//     PlcTask Outputs/GVL_iXlinker.Device_1_EtherCAT.Term_1_EK1200.Term_2_EL6002.COM_RxPDO_Map_Outputs_Channel_1.Data_Out[3] <-> COM RxPDO-Map Outputs Channel 1/Data Out 3
//     PlcTask Outputs/GVL_iXlinker.Device_1_EtherCAT.Term_1_EK1200.Term_2_EL6002.COM_RxPDO_Map_Outputs_Channel_1.Data_Out[4] <-> COM RxPDO-Map Outputs Channel 1/Data Out 4
//     PlcTask Outputs/GVL_iXlinker.Device_1_EtherCAT.Term_1_EK1200.Term_2_EL6002.COM_RxPDO_Map_Outputs_Channel_1.Data_Out[5] <-> COM RxPDO-Map Outputs Channel 1/Data Out 5
//     PlcTask Outputs/GVL_iXlinker.Device_1_EtherCAT.Term_1_EK1200.Term_2_EL6002.COM_RxPDO_Map_Outputs_Channel_1.Data_Out[6] <-> COM RxPDO-Map Outputs Channel 1/Data Out 6
//     PlcTask Outputs/GVL_iXlinker.Device_1_EtherCAT.Term_1_EK1200.Term_2_EL6002.COM_RxPDO_Map_Outputs_Channel_1.Data_Out[7] <-> COM RxPDO-Map Outputs Channel 1/Data Out 7
//     PlcTask Outputs/GVL_iXlinker.Device_1_EtherCAT.Term_1_EK1200.Term_2_EL6002.COM_RxPDO_Map_Outputs_Channel_1.Data_Out[8] <-> COM RxPDO-Map Outputs Channel 1/Data Out 8
//     PlcTask Outputs/GVL_iXlinker.Device_1_EtherCAT.Term_1_EK1200.Term_2_EL6002.COM_RxPDO_Map_Outputs_Channel_1.Data_Out[9] <-> COM RxPDO-Map Outputs Channel 1/Data Out 9
//     PlcTask Outputs/GVL_iXlinker.Device_1_EtherCAT.Term_1_EK1200.Term_2_EL6002.COM_RxPDO_Map_Outputs_Channel_2.Data_Out[0] <-> COM RxPDO-Map Outputs Channel 2/Data Out 0
//     PlcTask Outputs/GVL_iXlinker.Device_1_EtherCAT.Term_1_EK1200.Term_2_EL6002.COM_RxPDO_Map_Outputs_Channel_2.Data_Out[10] <-> COM RxPDO-Map Outputs Channel 2/Data Out 10
//     PlcTask Outputs/GVL_iXlinker.Device_1_EtherCAT.Term_1_EK1200.Term_2_EL6002.COM_RxPDO_Map_Outputs_Channel_2.Data_Out[11] <-> COM RxPDO-Map Outputs Channel 2/Data Out 11
//     PlcTask Outputs/GVL_iXlinker.Device_1_EtherCAT.Term_1_EK1200.Term_2_EL6002.COM_RxPDO_Map_Outputs_Channel_2.Data_Out[12] <-> COM RxPDO-Map Outputs Channel 2/Data Out 12
//     PlcTask Outputs/GVL_iXlinker.Device_1_EtherCAT.Term_1_EK1200.Term_2_EL6002.COM_RxPDO_Map_Outputs_Channel_2.Data_Out[13] <-> COM RxPDO-Map Outputs Channel 2/Data Out 13
//     PlcTask Outputs/GVL_iXlinker.Device_1_EtherCAT.Term_1_EK1200.Term_2_EL6002.COM_RxPDO_Map_Outputs_Channel_2.Data_Out[14] <-> COM RxPDO-Map Outputs Channel 2/Data Out 14
//     PlcTask Outputs/GVL_iXlinker.Device_1_EtherCAT.Term_1_EK1200.Term_2_EL6002.COM_RxPDO_Map_Outputs_Channel_2.Data_Out[15] <-> COM RxPDO-Map Outputs Channel 2/Data Out 15
//     PlcTask Outputs/GVL_iXlinker.Device_1_EtherCAT.Term_1_EK1200.Term_2_EL6002.COM_RxPDO_Map_Outputs_Channel_2.Data_Out[16] <-> COM RxPDO-Map Outputs Channel 2/Data Out 16
//     PlcTask Outputs/GVL_iXlinker.Device_1_EtherCAT.Term_1_EK1200.Term_2_EL6002.COM_RxPDO_Map_Outputs_Channel_2.Data_Out[17] <-> COM RxPDO-Map Outputs Channel 2/Data Out 17
//     PlcTask Outputs/GVL_iXlinker.Device_1_EtherCAT.Term_1_EK1200.Term_2_EL6002.COM_RxPDO_Map_Outputs_Channel_2.Data_Out[18] <-> COM RxPDO-Map Outputs Channel 2/Data Out 18
//     PlcTask Outputs/GVL_iXlinker.Device_1_EtherCAT.Term_1_EK1200.Term_2_EL6002.COM_RxPDO_Map_Outputs_Channel_2.Data_Out[19] <-> COM RxPDO-Map Outputs Channel 2/Data Out 19
//     PlcTask Outputs/GVL_iXlinker.Device_1_EtherCAT.Term_1_EK1200.Term_2_EL6002.COM_RxPDO_Map_Outputs_Channel_2.Data_Out[1] <-> COM RxPDO-Map Outputs Channel 2/Data Out 1
//     PlcTask Outputs/GVL_iXlinker.Device_1_EtherCAT.Term_1_EK1200.Term_2_EL6002.COM_RxPDO_Map_Outputs_Channel_2.Data_Out[20] <-> COM RxPDO-Map Outputs Channel 2/Data Out 20
//     PlcTask Outputs/GVL_iXlinker.Device_1_EtherCAT.Term_1_EK1200.Term_2_EL6002.COM_RxPDO_Map_Outputs_Channel_2.Data_Out[21] <-> COM RxPDO-Map Outputs Channel 2/Data Out 21
//     PlcTask Outputs/GVL_iXlinker.Device_1_EtherCAT.Term_1_EK1200.Term_2_EL6002.COM_RxPDO_Map_Outputs_Channel_2.Data_Out[2] <-> COM RxPDO-Map Outputs Channel 2/Data Out 2
//     PlcTask Outputs/GVL_iXlinker.Device_1_EtherCAT.Term_1_EK1200.Term_2_EL6002.COM_RxPDO_Map_Outputs_Channel_2.Data_Out[3] <-> COM RxPDO-Map Outputs Channel 2/Data Out 3
//     PlcTask Outputs/GVL_iXlinker.Device_1_EtherCAT.Term_1_EK1200.Term_2_EL6002.COM_RxPDO_Map_Outputs_Channel_2.Data_Out[4] <-> COM RxPDO-Map Outputs Channel 2/Data Out 4
//     PlcTask Outputs/GVL_iXlinker.Device_1_EtherCAT.Term_1_EK1200.Term_2_EL6002.COM_RxPDO_Map_Outputs_Channel_2.Data_Out[5] <-> COM RxPDO-Map Outputs Channel 2/Data Out 5
//     PlcTask Outputs/GVL_iXlinker.Device_1_EtherCAT.Term_1_EK1200.Term_2_EL6002.COM_RxPDO_Map_Outputs_Channel_2.Data_Out[6] <-> COM RxPDO-Map Outputs Channel 2/Data Out 6
//     PlcTask Outputs/GVL_iXlinker.Device_1_EtherCAT.Term_1_EK1200.Term_2_EL6002.COM_RxPDO_Map_Outputs_Channel_2.Data_Out[7] <-> COM RxPDO-Map Outputs Channel 2/Data Out 7
//     PlcTask Outputs/GVL_iXlinker.Device_1_EtherCAT.Term_1_EK1200.Term_2_EL6002.COM_RxPDO_Map_Outputs_Channel_2.Data_Out[8] <-> COM RxPDO-Map Outputs Channel 2/Data Out 8
//     PlcTask Outputs/GVL_iXlinker.Device_1_EtherCAT.Term_1_EK1200.Term_2_EL6002.COM_RxPDO_Map_Outputs_Channel_2.Data_Out[9] <-> COM RxPDO-Map Outputs Channel 2/Data Out 9
//   TcoIoTests/TcoIoTests Instance <-> Device 1 (EtherCAT)/Term 1 (EK1200)/Term 3 (EL1809)
//     PlcTask Inputs/GVL_iXlinker.Device_1_EtherCAT.Term_1_EK1200.Term_3_EL1809.Channel_{1..16}.Input <-> Channel {1..16}/Input  (16 links)
//     PlcTask Inputs/GVL_iXlinker.Device_1_EtherCAT.Term_1_EK1200.Term_3_EL1809.InfoData.State <-> InfoData/State
//     PlcTask Inputs/GVL_iXlinker.Device_1_EtherCAT.Term_1_EK1200.Term_3_EL1809.WcState.InputToggle <-> WcState/InputToggle
//     PlcTask Inputs/GVL_iXlinker.Device_1_EtherCAT.Term_1_EK1200.Term_3_EL1809.WcState.WcState <-> WcState/WcState
//   TcoIoTests/TcoIoTests Instance <-> Device 1 (EtherCAT)/Term 1 (EK1200)/Term 4 (EL2809)
//     PlcTask Inputs/GVL_iXlinker.Device_1_EtherCAT.Term_1_EK1200.Term_4_EL2809.InfoData.State <-> InfoData/State
//     PlcTask Inputs/GVL_iXlinker.Device_1_EtherCAT.Term_1_EK1200.Term_4_EL2809.WcState.WcState <-> WcState/WcState
//     PlcTask Outputs/GVL_iXlinker.Device_1_EtherCAT.Term_1_EK1200.Term_4_EL2809.Channel_{1..16}.Output <-> Channel {1..16}/Output  (16 links)
//   TcoIoTests/TcoIoTests Instance <-> Device 1 (EtherCAT)/Term 1 (EK1200)/Term 5 (EL4004)
//     PlcTask Inputs/GVL_iXlinker.Device_1_EtherCAT.Term_1_EK1200.Term_5_EL4004.InfoData.AdsAddr <-> InfoData/AdsAddr
//     PlcTask Inputs/GVL_iXlinker.Device_1_EtherCAT.Term_1_EK1200.Term_5_EL4004.InfoData.State <-> InfoData/State
//     PlcTask Inputs/GVL_iXlinker.Device_1_EtherCAT.Term_1_EK1200.Term_5_EL4004.WcState.WcState <-> WcState/WcState
//     PlcTask Outputs/GVL_iXlinker.Device_1_EtherCAT.Term_1_EK1200.Term_5_EL4004.AO_Outputs_Channel_{1..4}.Analog_output <-> AO Outputs Channel {1..4}/Analog output  (4 links)
//   TcoIoTests/TcoIoTests Instance <-> Device 1 (EtherCAT)/Term 1 (EK1200)/Term 6 (EL2809)
//     PlcTask Inputs/GVL_iXlinker.Device_1_EtherCAT.Term_1_EK1200.Term_6_EL2809.InfoData.State <-> InfoData/State
//     PlcTask Inputs/GVL_iXlinker.Device_1_EtherCAT.Term_1_EK1200.Term_6_EL2809.WcState.WcState <-> WcState/WcState
//     PlcTask Outputs/GVL_iXlinker.Device_1_EtherCAT.Term_1_EK1200.Term_6_EL2809.Channel_{1..16}.Output <-> Channel {1..16}/Output  (16 links)
//   TcoIoTests/TcoIoTests Instance <-> Device 1 (EtherCAT)/Term 1 (EK1200)/Term 7 (EL6001)
//     PlcTask Inputs/GVL_iXlinker.Device_1_EtherCAT.Term_1_EK1200.Term_7_EL6001.COM_Inputs.Data_In[{0..21}] <-> COM Inputs/Data In {0..21}  (22 links)
//     PlcTask Inputs/GVL_iXlinker.Device_1_EtherCAT.Term_1_EK1200.Term_7_EL6001.COM_Inputs.Status/Buffer_full <-> COM Inputs/Status/Buffer full
//     PlcTask Inputs/GVL_iXlinker.Device_1_EtherCAT.Term_1_EK1200.Term_7_EL6001.COM_Inputs.Status/Framing_error <-> COM Inputs/Status/Framing error
//     PlcTask Inputs/GVL_iXlinker.Device_1_EtherCAT.Term_1_EK1200.Term_7_EL6001.COM_Inputs.Status/Init_accepted <-> COM Inputs/Status/Init accepted
//     PlcTask Inputs/GVL_iXlinker.Device_1_EtherCAT.Term_1_EK1200.Term_7_EL6001.COM_Inputs.Status/Input_length <-> COM Inputs/Status/Input length
//     PlcTask Inputs/GVL_iXlinker.Device_1_EtherCAT.Term_1_EK1200.Term_7_EL6001.COM_Inputs.Status/Overrun_error <-> COM Inputs/Status/Overrun error
//     PlcTask Inputs/GVL_iXlinker.Device_1_EtherCAT.Term_1_EK1200.Term_7_EL6001.COM_Inputs.Status/Parity_error <-> COM Inputs/Status/Parity error
//     PlcTask Inputs/GVL_iXlinker.Device_1_EtherCAT.Term_1_EK1200.Term_7_EL6001.COM_Inputs.Status/Receive_request <-> COM Inputs/Status/Receive request
//     PlcTask Inputs/GVL_iXlinker.Device_1_EtherCAT.Term_1_EK1200.Term_7_EL6001.COM_Inputs.Status/Transmit_accepted <-> COM Inputs/Status/Transmit accepted
//     PlcTask Inputs/GVL_iXlinker.Device_1_EtherCAT.Term_1_EK1200.Term_7_EL6001.InfoData.AdsAddr <-> InfoData/AdsAddr
//     PlcTask Inputs/GVL_iXlinker.Device_1_EtherCAT.Term_1_EK1200.Term_7_EL6001.InfoData.State <-> InfoData/State
//     PlcTask Inputs/GVL_iXlinker.Device_1_EtherCAT.Term_1_EK1200.Term_7_EL6001.WcState.InputToggle <-> WcState/InputToggle
//     PlcTask Inputs/GVL_iXlinker.Device_1_EtherCAT.Term_1_EK1200.Term_7_EL6001.WcState.WcState <-> WcState/WcState
//     PlcTask Outputs/GVL_iXlinker.Device_1_EtherCAT.Term_1_EK1200.Term_7_EL6001.COM_Outputs.Ctrl/Init_request <-> COM Outputs/Ctrl/Init request
//     PlcTask Outputs/GVL_iXlinker.Device_1_EtherCAT.Term_1_EK1200.Term_7_EL6001.COM_Outputs.Ctrl/Output_length <-> COM Outputs/Ctrl/Output length
//     PlcTask Outputs/GVL_iXlinker.Device_1_EtherCAT.Term_1_EK1200.Term_7_EL6001.COM_Outputs.Ctrl/Receive_accepted <-> COM Outputs/Ctrl/Receive accepted
//     PlcTask Outputs/GVL_iXlinker.Device_1_EtherCAT.Term_1_EK1200.Term_7_EL6001.COM_Outputs.Ctrl/Send_continues <-> COM Outputs/Ctrl/Send continues
//     PlcTask Outputs/GVL_iXlinker.Device_1_EtherCAT.Term_1_EK1200.Term_7_EL6001.COM_Outputs.Ctrl/Transmit_request <-> COM Outputs/Ctrl/Transmit request
//     PlcTask Outputs/GVL_iXlinker.Device_1_EtherCAT.Term_1_EK1200.Term_7_EL6001.COM_Outputs.Data_Out[{0..21}] <-> COM Outputs/Data Out {0..21}  (22 links)
//   TcoIoTests/TcoIoTests Instance <-> Device 2 (EtherCAT)
//     PlcTask Inputs/GVL_iXlinker.Device_2_EtherCAT.InfoData.AmsNetId <-> InfoData/AmsNetId
//     PlcTask Inputs/GVL_iXlinker.Device_2_EtherCAT.InfoData.CfgSlaveCount <-> InfoData/CfgSlaveCount
//     PlcTask Inputs/GVL_iXlinker.Device_2_EtherCAT.InfoData.ChangeCount <-> InfoData/ChangeCount
//     PlcTask Inputs/GVL_iXlinker.Device_2_EtherCAT.InfoData.DevId <-> InfoData/DevId
//     PlcTask Inputs/GVL_iXlinker.Device_2_EtherCAT.Inputs.DevState <-> Inputs/DevState
//     PlcTask Inputs/GVL_iXlinker.Device_2_EtherCAT.Inputs.Frm0InputToggle <-> Inputs/Frm0InputToggle
//     PlcTask Inputs/GVL_iXlinker.Device_2_EtherCAT.Inputs.Frm0State <-> Inputs/Frm0State
//     PlcTask Inputs/GVL_iXlinker.Device_2_EtherCAT.Inputs.Frm0WcState <-> Inputs/Frm0WcState
//     PlcTask Inputs/GVL_iXlinker.Device_2_EtherCAT.Inputs.SlaveCount <-> Inputs/SlaveCount
//     PlcTask Outputs/GVL_iXlinker.Device_2_EtherCAT.Outputs.DevCtrl <-> Outputs/DevCtrl
//     PlcTask Outputs/GVL_iXlinker.Device_2_EtherCAT.Outputs.Frm0Ctrl <-> Outputs/Frm0Ctrl
//     PlcTask Outputs/GVL_iXlinker.Device_2_EtherCAT.Outputs.Frm0WcCtrl <-> Outputs/Frm0WcCtrl
//   TcoIoTests/TcoIoTests Instance <-> Device 2 (EtherCAT)/Term 9 (EK1100)
//     PlcTask Inputs/GVL_iXlinker.Device_2_EtherCAT.Term_9_EK1100.InfoData.State <-> InfoData/State
//   TcoIoTests/TcoIoTests Instance <-> Device 2 (EtherCAT)/Term 9 (EK1100)/Term 10 (EK1122)
//     PlcTask Inputs/GVL_iXlinker.Device_2_EtherCAT.Term_9_EK1100.Term_10_EK1122.InfoData.State <-> InfoData/State
//   TcoIoTests/TcoIoTests Instance <-> Device 2 (EtherCAT)/Term 9 (EK1100)/Term 10 (EK1122)/Term 11 (EK1100)
//     PlcTask Inputs/GVL_iXlinker.Device_2_EtherCAT.Term_9_EK1100.Term_10_EK1122.Term_11_EK1100.InfoData.State <-> InfoData/State
//   TcoIoTests/TcoIoTests Instance <-> Device 2 (EtherCAT)/Term 9 (EK1100)/Term 10 (EK1122)/Term 11 (EK1100)/Term 12 (EL3174-0002)
//     PlcTask Inputs/GVL_iXlinker.Device_2_EtherCAT.Term_9_EK1100.Term_10_EK1122.Term_11_EK1100.Term_12_EL3174_0002.AI_Standard_Channel_1.Status/Error <-> AI Standard Channel 1/Status/Error
//     PlcTask Inputs/GVL_iXlinker.Device_2_EtherCAT.Term_9_EK1100.Term_10_EK1122.Term_11_EK1100.Term_12_EL3174_0002.AI_Standard_Channel_2.Status/Error <-> AI Standard Channel 2/Status/Error
//     PlcTask Inputs/GVL_iXlinker.Device_2_EtherCAT.Term_9_EK1100.Term_10_EK1122.Term_11_EK1100.Term_12_EL3174_0002.AI_Standard_Channel_3.Status/Error <-> AI Standard Channel 3/Status/Error
//     PlcTask Inputs/GVL_iXlinker.Device_2_EtherCAT.Term_9_EK1100.Term_10_EK1122.Term_11_EK1100.Term_12_EL3174_0002.AI_Standard_Channel_4.Status/Error <-> AI Standard Channel 4/Status/Error
//     PlcTask Inputs/GVL_iXlinker.Device_2_EtherCAT.Term_9_EK1100.Term_10_EK1122.Term_11_EK1100.Term_12_EL3174_0002.AI_Standard_Channel_1.Status/Limit_1 <-> AI Standard Channel 1/Status/Limit 1
//     PlcTask Inputs/GVL_iXlinker.Device_2_EtherCAT.Term_9_EK1100.Term_10_EK1122.Term_11_EK1100.Term_12_EL3174_0002.AI_Standard_Channel_1.Status/Limit_2 <-> AI Standard Channel 1/Status/Limit 2
//     PlcTask Inputs/GVL_iXlinker.Device_2_EtherCAT.Term_9_EK1100.Term_10_EK1122.Term_11_EK1100.Term_12_EL3174_0002.AI_Standard_Channel_2.Status/Limit_1 <-> AI Standard Channel 2/Status/Limit 1
//     PlcTask Inputs/GVL_iXlinker.Device_2_EtherCAT.Term_9_EK1100.Term_10_EK1122.Term_11_EK1100.Term_12_EL3174_0002.AI_Standard_Channel_2.Status/Limit_2 <-> AI Standard Channel 2/Status/Limit 2
//     PlcTask Inputs/GVL_iXlinker.Device_2_EtherCAT.Term_9_EK1100.Term_10_EK1122.Term_11_EK1100.Term_12_EL3174_0002.AI_Standard_Channel_3.Status/Limit_1 <-> AI Standard Channel 3/Status/Limit 1
//     PlcTask Inputs/GVL_iXlinker.Device_2_EtherCAT.Term_9_EK1100.Term_10_EK1122.Term_11_EK1100.Term_12_EL3174_0002.AI_Standard_Channel_3.Status/Limit_2 <-> AI Standard Channel 3/Status/Limit 2
//     PlcTask Inputs/GVL_iXlinker.Device_2_EtherCAT.Term_9_EK1100.Term_10_EK1122.Term_11_EK1100.Term_12_EL3174_0002.AI_Standard_Channel_4.Status/Limit_1 <-> AI Standard Channel 4/Status/Limit 1
//     PlcTask Inputs/GVL_iXlinker.Device_2_EtherCAT.Term_9_EK1100.Term_10_EK1122.Term_11_EK1100.Term_12_EL3174_0002.AI_Standard_Channel_4.Status/Limit_2 <-> AI Standard Channel 4/Status/Limit 2
//     PlcTask Inputs/GVL_iXlinker.Device_2_EtherCAT.Term_9_EK1100.Term_10_EK1122.Term_11_EK1100.Term_12_EL3174_0002.AI_Standard_Channel_1.Status/Overrange <-> AI Standard Channel 1/Status/Overrange
//     PlcTask Inputs/GVL_iXlinker.Device_2_EtherCAT.Term_9_EK1100.Term_10_EK1122.Term_11_EK1100.Term_12_EL3174_0002.AI_Standard_Channel_2.Status/Overrange <-> AI Standard Channel 2/Status/Overrange
//     PlcTask Inputs/GVL_iXlinker.Device_2_EtherCAT.Term_9_EK1100.Term_10_EK1122.Term_11_EK1100.Term_12_EL3174_0002.AI_Standard_Channel_3.Status/Overrange <-> AI Standard Channel 3/Status/Overrange
//     PlcTask Inputs/GVL_iXlinker.Device_2_EtherCAT.Term_9_EK1100.Term_10_EK1122.Term_11_EK1100.Term_12_EL3174_0002.AI_Standard_Channel_4.Status/Overrange <-> AI Standard Channel 4/Status/Overrange
//     PlcTask Inputs/GVL_iXlinker.Device_2_EtherCAT.Term_9_EK1100.Term_10_EK1122.Term_11_EK1100.Term_12_EL3174_0002.AI_Standard_Channel_1.Status/Sync_error <-> AI Standard Channel 1/Status/Sync error
//     PlcTask Inputs/GVL_iXlinker.Device_2_EtherCAT.Term_9_EK1100.Term_10_EK1122.Term_11_EK1100.Term_12_EL3174_0002.AI_Standard_Channel_2.Status/Sync_error <-> AI Standard Channel 2/Status/Sync error
//     PlcTask Inputs/GVL_iXlinker.Device_2_EtherCAT.Term_9_EK1100.Term_10_EK1122.Term_11_EK1100.Term_12_EL3174_0002.AI_Standard_Channel_3.Status/Sync_error <-> AI Standard Channel 3/Status/Sync error
//     PlcTask Inputs/GVL_iXlinker.Device_2_EtherCAT.Term_9_EK1100.Term_10_EK1122.Term_11_EK1100.Term_12_EL3174_0002.AI_Standard_Channel_4.Status/Sync_error <-> AI Standard Channel 4/Status/Sync error
//     PlcTask Inputs/GVL_iXlinker.Device_2_EtherCAT.Term_9_EK1100.Term_10_EK1122.Term_11_EK1100.Term_12_EL3174_0002.AI_Standard_Channel_1.Status/TxPDO_State <-> AI Standard Channel 1/Status/TxPDO State
//     PlcTask Inputs/GVL_iXlinker.Device_2_EtherCAT.Term_9_EK1100.Term_10_EK1122.Term_11_EK1100.Term_12_EL3174_0002.AI_Standard_Channel_2.Status/TxPDO_State <-> AI Standard Channel 2/Status/TxPDO State
//     PlcTask Inputs/GVL_iXlinker.Device_2_EtherCAT.Term_9_EK1100.Term_10_EK1122.Term_11_EK1100.Term_12_EL3174_0002.AI_Standard_Channel_3.Status/TxPDO_State <-> AI Standard Channel 3/Status/TxPDO State
//     PlcTask Inputs/GVL_iXlinker.Device_2_EtherCAT.Term_9_EK1100.Term_10_EK1122.Term_11_EK1100.Term_12_EL3174_0002.AI_Standard_Channel_4.Status/TxPDO_State <-> AI Standard Channel 4/Status/TxPDO State
//     PlcTask Inputs/GVL_iXlinker.Device_2_EtherCAT.Term_9_EK1100.Term_10_EK1122.Term_11_EK1100.Term_12_EL3174_0002.AI_Standard_Channel_1.Status/TxPDO_Toggle <-> AI Standard Channel 1/Status/TxPDO Toggle
//     PlcTask Inputs/GVL_iXlinker.Device_2_EtherCAT.Term_9_EK1100.Term_10_EK1122.Term_11_EK1100.Term_12_EL3174_0002.AI_Standard_Channel_2.Status/TxPDO_Toggle <-> AI Standard Channel 2/Status/TxPDO Toggle
//     PlcTask Inputs/GVL_iXlinker.Device_2_EtherCAT.Term_9_EK1100.Term_10_EK1122.Term_11_EK1100.Term_12_EL3174_0002.AI_Standard_Channel_3.Status/TxPDO_Toggle <-> AI Standard Channel 3/Status/TxPDO Toggle
//     PlcTask Inputs/GVL_iXlinker.Device_2_EtherCAT.Term_9_EK1100.Term_10_EK1122.Term_11_EK1100.Term_12_EL3174_0002.AI_Standard_Channel_4.Status/TxPDO_Toggle <-> AI Standard Channel 4/Status/TxPDO Toggle
//     PlcTask Inputs/GVL_iXlinker.Device_2_EtherCAT.Term_9_EK1100.Term_10_EK1122.Term_11_EK1100.Term_12_EL3174_0002.AI_Standard_Channel_1.Status/Underrange <-> AI Standard Channel 1/Status/Underrange
//     PlcTask Inputs/GVL_iXlinker.Device_2_EtherCAT.Term_9_EK1100.Term_10_EK1122.Term_11_EK1100.Term_12_EL3174_0002.AI_Standard_Channel_2.Status/Underrange <-> AI Standard Channel 2/Status/Underrange
//     PlcTask Inputs/GVL_iXlinker.Device_2_EtherCAT.Term_9_EK1100.Term_10_EK1122.Term_11_EK1100.Term_12_EL3174_0002.AI_Standard_Channel_3.Status/Underrange <-> AI Standard Channel 3/Status/Underrange
//     PlcTask Inputs/GVL_iXlinker.Device_2_EtherCAT.Term_9_EK1100.Term_10_EK1122.Term_11_EK1100.Term_12_EL3174_0002.AI_Standard_Channel_4.Status/Underrange <-> AI Standard Channel 4/Status/Underrange
//     PlcTask Inputs/GVL_iXlinker.Device_2_EtherCAT.Term_9_EK1100.Term_10_EK1122.Term_11_EK1100.Term_12_EL3174_0002.AI_Standard_Channel_1.Value <-> AI Standard Channel 1/Value
//     PlcTask Inputs/GVL_iXlinker.Device_2_EtherCAT.Term_9_EK1100.Term_10_EK1122.Term_11_EK1100.Term_12_EL3174_0002.AI_Standard_Channel_2.Value <-> AI Standard Channel 2/Value
//     PlcTask Inputs/GVL_iXlinker.Device_2_EtherCAT.Term_9_EK1100.Term_10_EK1122.Term_11_EK1100.Term_12_EL3174_0002.AI_Standard_Channel_3.Value <-> AI Standard Channel 3/Value
//     PlcTask Inputs/GVL_iXlinker.Device_2_EtherCAT.Term_9_EK1100.Term_10_EK1122.Term_11_EK1100.Term_12_EL3174_0002.AI_Standard_Channel_4.Value <-> AI Standard Channel 4/Value
//     PlcTask Inputs/GVL_iXlinker.Device_2_EtherCAT.Term_9_EK1100.Term_10_EK1122.Term_11_EK1100.Term_12_EL3174_0002.InfoData.AdsAddr <-> InfoData/AdsAddr
//     PlcTask Inputs/GVL_iXlinker.Device_2_EtherCAT.Term_9_EK1100.Term_10_EK1122.Term_11_EK1100.Term_12_EL3174_0002.InfoData.State <-> InfoData/State
//     PlcTask Inputs/GVL_iXlinker.Device_2_EtherCAT.Term_9_EK1100.Term_10_EK1122.Term_11_EK1100.Term_12_EL3174_0002.WcState.InputToggle <-> WcState/InputToggle
//     PlcTask Inputs/GVL_iXlinker.Device_2_EtherCAT.Term_9_EK1100.Term_10_EK1122.Term_11_EK1100.Term_12_EL3174_0002.WcState.WcState <-> WcState/WcState
//   TcoIoTests/TcoIoTests Instance <-> Device 2 (EtherCAT)/Term 9 (EK1100)/Term 10 (EK1122)/Term 11 (EK1100)/Term 13 (EL6001)
//     PlcTask Inputs/GVL_iXlinker.Device_2_EtherCAT.Term_9_EK1100.Term_10_EK1122.Term_11_EK1100.Term_13_EL6001.COM_Inputs.Data_In[{0..21}] <-> COM Inputs/Data In {0..21}  (22 links)
//     PlcTask Inputs/GVL_iXlinker.Device_2_EtherCAT.Term_9_EK1100.Term_10_EK1122.Term_11_EK1100.Term_13_EL6001.COM_Inputs.Status/Buffer_full <-> COM Inputs/Status/Buffer full
//     PlcTask Inputs/GVL_iXlinker.Device_2_EtherCAT.Term_9_EK1100.Term_10_EK1122.Term_11_EK1100.Term_13_EL6001.COM_Inputs.Status/Framing_error <-> COM Inputs/Status/Framing error
//     PlcTask Inputs/GVL_iXlinker.Device_2_EtherCAT.Term_9_EK1100.Term_10_EK1122.Term_11_EK1100.Term_13_EL6001.COM_Inputs.Status/Init_accepted <-> COM Inputs/Status/Init accepted
//     PlcTask Inputs/GVL_iXlinker.Device_2_EtherCAT.Term_9_EK1100.Term_10_EK1122.Term_11_EK1100.Term_13_EL6001.COM_Inputs.Status/Input_length <-> COM Inputs/Status/Input length
//     PlcTask Inputs/GVL_iXlinker.Device_2_EtherCAT.Term_9_EK1100.Term_10_EK1122.Term_11_EK1100.Term_13_EL6001.COM_Inputs.Status/Overrun_error <-> COM Inputs/Status/Overrun error
//     PlcTask Inputs/GVL_iXlinker.Device_2_EtherCAT.Term_9_EK1100.Term_10_EK1122.Term_11_EK1100.Term_13_EL6001.COM_Inputs.Status/Parity_error <-> COM Inputs/Status/Parity error
//     PlcTask Inputs/GVL_iXlinker.Device_2_EtherCAT.Term_9_EK1100.Term_10_EK1122.Term_11_EK1100.Term_13_EL6001.COM_Inputs.Status/Receive_request <-> COM Inputs/Status/Receive request
//     PlcTask Inputs/GVL_iXlinker.Device_2_EtherCAT.Term_9_EK1100.Term_10_EK1122.Term_11_EK1100.Term_13_EL6001.COM_Inputs.Status/Transmit_accepted <-> COM Inputs/Status/Transmit accepted
//     PlcTask Inputs/GVL_iXlinker.Device_2_EtherCAT.Term_9_EK1100.Term_10_EK1122.Term_11_EK1100.Term_13_EL6001.InfoData.AdsAddr <-> InfoData/AdsAddr
//     PlcTask Inputs/GVL_iXlinker.Device_2_EtherCAT.Term_9_EK1100.Term_10_EK1122.Term_11_EK1100.Term_13_EL6001.InfoData.State <-> InfoData/State
//     PlcTask Inputs/GVL_iXlinker.Device_2_EtherCAT.Term_9_EK1100.Term_10_EK1122.Term_11_EK1100.Term_13_EL6001.WcState.InputToggle <-> WcState/InputToggle
//     PlcTask Inputs/GVL_iXlinker.Device_2_EtherCAT.Term_9_EK1100.Term_10_EK1122.Term_11_EK1100.Term_13_EL6001.WcState.WcState <-> WcState/WcState
//     PlcTask Outputs/GVL_iXlinker.Device_2_EtherCAT.Term_9_EK1100.Term_10_EK1122.Term_11_EK1100.Term_13_EL6001.COM_Outputs.Ctrl/Init_request <-> COM Outputs/Ctrl/Init request
//     PlcTask Outputs/GVL_iXlinker.Device_2_EtherCAT.Term_9_EK1100.Term_10_EK1122.Term_11_EK1100.Term_13_EL6001.COM_Outputs.Ctrl/Output_length <-> COM Outputs/Ctrl/Output length
//     PlcTask Outputs/GVL_iXlinker.Device_2_EtherCAT.Term_9_EK1100.Term_10_EK1122.Term_11_EK1100.Term_13_EL6001.COM_Outputs.Ctrl/Receive_accepted <-> COM Outputs/Ctrl/Receive accepted
//     PlcTask Outputs/GVL_iXlinker.Device_2_EtherCAT.Term_9_EK1100.Term_10_EK1122.Term_11_EK1100.Term_13_EL6001.COM_Outputs.Ctrl/Send_continues <-> COM Outputs/Ctrl/Send continues
//     PlcTask Outputs/GVL_iXlinker.Device_2_EtherCAT.Term_9_EK1100.Term_10_EK1122.Term_11_EK1100.Term_13_EL6001.COM_Outputs.Ctrl/Transmit_request <-> COM Outputs/Ctrl/Transmit request
//     PlcTask Outputs/GVL_iXlinker.Device_2_EtherCAT.Term_9_EK1100.Term_10_EK1122.Term_11_EK1100.Term_13_EL6001.COM_Outputs.Data_Out[{0..21}] <-> COM Outputs/Data Out {0..21}  (22 links)
//   TcoIoTests/TcoIoTests Instance <-> Device 2 (EtherCAT)/Term 9 (EK1100)/Term 10 (EK1122)/Term 11 (EK1100)/Term 14 (EL3011)
//     PlcTask Inputs/GVL_iXlinker.Device_2_EtherCAT.Term_9_EK1100.Term_10_EK1122.Term_11_EK1100.Term_14_EL3011.AI_Standard.Status/Error <-> AI Standard/Status/Error
//     PlcTask Inputs/GVL_iXlinker.Device_2_EtherCAT.Term_9_EK1100.Term_10_EK1122.Term_11_EK1100.Term_14_EL3011.AI_Standard.Status/Limit_1 <-> AI Standard/Status/Limit 1
//     PlcTask Inputs/GVL_iXlinker.Device_2_EtherCAT.Term_9_EK1100.Term_10_EK1122.Term_11_EK1100.Term_14_EL3011.AI_Standard.Status/Limit_2 <-> AI Standard/Status/Limit 2
//     PlcTask Inputs/GVL_iXlinker.Device_2_EtherCAT.Term_9_EK1100.Term_10_EK1122.Term_11_EK1100.Term_14_EL3011.AI_Standard.Status/Overrange <-> AI Standard/Status/Overrange
//     PlcTask Inputs/GVL_iXlinker.Device_2_EtherCAT.Term_9_EK1100.Term_10_EK1122.Term_11_EK1100.Term_14_EL3011.AI_Standard.Status/TxPDO_State <-> AI Standard/Status/TxPDO State
//     PlcTask Inputs/GVL_iXlinker.Device_2_EtherCAT.Term_9_EK1100.Term_10_EK1122.Term_11_EK1100.Term_14_EL3011.AI_Standard.Status/TxPDO_Toggle <-> AI Standard/Status/TxPDO Toggle
//     PlcTask Inputs/GVL_iXlinker.Device_2_EtherCAT.Term_9_EK1100.Term_10_EK1122.Term_11_EK1100.Term_14_EL3011.AI_Standard.Status/Underrange <-> AI Standard/Status/Underrange
//     PlcTask Inputs/GVL_iXlinker.Device_2_EtherCAT.Term_9_EK1100.Term_10_EK1122.Term_11_EK1100.Term_14_EL3011.AI_Standard.Value <-> AI Standard/Value
//     PlcTask Inputs/GVL_iXlinker.Device_2_EtherCAT.Term_9_EK1100.Term_10_EK1122.Term_11_EK1100.Term_14_EL3011.InfoData.AdsAddr <-> InfoData/AdsAddr
//     PlcTask Inputs/GVL_iXlinker.Device_2_EtherCAT.Term_9_EK1100.Term_10_EK1122.Term_11_EK1100.Term_14_EL3011.InfoData.State <-> InfoData/State
//     PlcTask Inputs/GVL_iXlinker.Device_2_EtherCAT.Term_9_EK1100.Term_10_EK1122.Term_11_EK1100.Term_14_EL3011.WcState.InputToggle <-> WcState/InputToggle
//     PlcTask Inputs/GVL_iXlinker.Device_2_EtherCAT.Term_9_EK1100.Term_10_EK1122.Term_11_EK1100.Term_14_EL3011.WcState.WcState <-> WcState/WcState
//   TcoIoTests/TcoIoTests Instance <-> Device 2 (EtherCAT)/Term 9 (EK1100)/Term 10 (EK1122)/Term 11 (EK1100)/Term 15 (EL2008)
//     PlcTask Inputs/GVL_iXlinker.Device_2_EtherCAT.Term_9_EK1100.Term_10_EK1122.Term_11_EK1100.Term_15_EL2008.InfoData.State <-> InfoData/State
//     PlcTask Inputs/GVL_iXlinker.Device_2_EtherCAT.Term_9_EK1100.Term_10_EK1122.Term_11_EK1100.Term_15_EL2008.WcState.WcState <-> WcState/WcState
//     PlcTask Outputs/GVL_iXlinker.Device_2_EtherCAT.Term_9_EK1100.Term_10_EK1122.Term_11_EK1100.Term_15_EL2008.Channel_{1..8}.Output <-> Channel {1..8}/Output  (8 links)
//   TcoIoTests/TcoIoTests Instance <-> Device 2 (EtherCAT)/Term 9 (EK1100)/Term 10 (EK1122)/Term 11 (EK1100)/Term 16 (EL2008)
//     PlcTask Inputs/GVL_iXlinker.Device_2_EtherCAT.Term_9_EK1100.Term_10_EK1122.Term_11_EK1100.Term_16_EL2008.InfoData.State <-> InfoData/State
//     PlcTask Inputs/GVL_iXlinker.Device_2_EtherCAT.Term_9_EK1100.Term_10_EK1122.Term_11_EK1100.Term_16_EL2008.WcState.WcState <-> WcState/WcState
//     PlcTask Outputs/GVL_iXlinker.Device_2_EtherCAT.Term_9_EK1100.Term_10_EK1122.Term_11_EK1100.Term_16_EL2008.Channel_{1..8}.Output <-> Channel {1..8}/Output  (8 links)
//   TcoIoTests/TcoIoTests Instance <-> Device 2 (EtherCAT)/Term 9 (EK1100)/Term 10 (EK1122)/Term 11 (EK1100)/Term 17 (EK1110)
//     PlcTask Inputs/GVL_iXlinker.Device_2_EtherCAT.Term_9_EK1100.Term_10_EK1122.Term_11_EK1100.Term_17_EK1110.InfoData.State <-> InfoData/State
//   TcoIoTests/TcoIoTests Instance <-> Device 2 (EtherCAT)/Term 9 (EK1100)/Term 10 (EK1122)/Term 18 (EK1100)
//     PlcTask Inputs/GVL_iXlinker.Device_2_EtherCAT.Term_9_EK1100.Term_10_EK1122.Term_18_EK1100.InfoData.State <-> InfoData/State
//   TcoIoTests/TcoIoTests Instance <-> Device 2 (EtherCAT)/Term 9 (EK1100)/Term 10 (EK1122)/Term 18 (EK1100)/Term 19 (EL1809)
//     PlcTask Inputs/GVL_iXlinker.Device_2_EtherCAT.Term_9_EK1100.Term_10_EK1122.Term_18_EK1100.Term_19_EL1809.Channel_{1..16}.Input <-> Channel {1..16}/Input  (16 links)
//     PlcTask Inputs/GVL_iXlinker.Device_2_EtherCAT.Term_9_EK1100.Term_10_EK1122.Term_18_EK1100.Term_19_EL1809.InfoData.State <-> InfoData/State
//     PlcTask Inputs/GVL_iXlinker.Device_2_EtherCAT.Term_9_EK1100.Term_10_EK1122.Term_18_EK1100.Term_19_EL1809.WcState.InputToggle <-> WcState/InputToggle
//     PlcTask Inputs/GVL_iXlinker.Device_2_EtherCAT.Term_9_EK1100.Term_10_EK1122.Term_18_EK1100.Term_19_EL1809.WcState.WcState <-> WcState/WcState
//   TcoIoTests/TcoIoTests Instance <-> Device 2 (EtherCAT)/Term 9 (EK1100)/Term 10 (EK1122)/Term 18 (EK1100)/Term 20 (EL2809)
//     PlcTask Inputs/GVL_iXlinker.Device_2_EtherCAT.Term_9_EK1100.Term_10_EK1122.Term_18_EK1100.Term_20_EL2809.InfoData.State <-> InfoData/State
//     PlcTask Inputs/GVL_iXlinker.Device_2_EtherCAT.Term_9_EK1100.Term_10_EK1122.Term_18_EK1100.Term_20_EL2809.WcState.WcState <-> WcState/WcState
//     PlcTask Outputs/GVL_iXlinker.Device_2_EtherCAT.Term_9_EK1100.Term_10_EK1122.Term_18_EK1100.Term_20_EL2809.Channel_{1..16}.Output <-> Channel {1..16}/Output  (16 links)
//   TcoIoTests/TcoIoTests Instance <-> Device 2 (EtherCAT)/Term 9 (EK1100)/Term 10 (EK1122)/Term 18 (EK1100)/Term 21 (EL1809)
//     PlcTask Inputs/GVL_iXlinker.Device_2_EtherCAT.Term_9_EK1100.Term_10_EK1122.Term_18_EK1100.Term_21_EL1809.Channel_{1..16}.Input <-> Channel {1..16}/Input  (16 links)
//     PlcTask Inputs/GVL_iXlinker.Device_2_EtherCAT.Term_9_EK1100.Term_10_EK1122.Term_18_EK1100.Term_21_EL1809.InfoData.State <-> InfoData/State
//     PlcTask Inputs/GVL_iXlinker.Device_2_EtherCAT.Term_9_EK1100.Term_10_EK1122.Term_18_EK1100.Term_21_EL1809.WcState.InputToggle <-> WcState/InputToggle
//     PlcTask Inputs/GVL_iXlinker.Device_2_EtherCAT.Term_9_EK1100.Term_10_EK1122.Term_18_EK1100.Term_21_EL1809.WcState.WcState <-> WcState/WcState
//   TcoIoTests/TcoIoTests Instance <-> Device 2 (EtherCAT)/Term 9 (EK1100)/Term 10 (EK1122)/Term 18 (EK1100)/Term 22 (EL3011)
//     PlcTask Inputs/GVL_iXlinker.Device_2_EtherCAT.Term_9_EK1100.Term_10_EK1122.Term_18_EK1100.Term_22_EL3011.AI_Standard.Status/Error <-> AI Standard/Status/Error
//     PlcTask Inputs/GVL_iXlinker.Device_2_EtherCAT.Term_9_EK1100.Term_10_EK1122.Term_18_EK1100.Term_22_EL3011.AI_Standard.Status/Limit_1 <-> AI Standard/Status/Limit 1
//     PlcTask Inputs/GVL_iXlinker.Device_2_EtherCAT.Term_9_EK1100.Term_10_EK1122.Term_18_EK1100.Term_22_EL3011.AI_Standard.Status/Limit_2 <-> AI Standard/Status/Limit 2
//     PlcTask Inputs/GVL_iXlinker.Device_2_EtherCAT.Term_9_EK1100.Term_10_EK1122.Term_18_EK1100.Term_22_EL3011.AI_Standard.Status/Overrange <-> AI Standard/Status/Overrange
//     PlcTask Inputs/GVL_iXlinker.Device_2_EtherCAT.Term_9_EK1100.Term_10_EK1122.Term_18_EK1100.Term_22_EL3011.AI_Standard.Status/TxPDO_State <-> AI Standard/Status/TxPDO State
//     PlcTask Inputs/GVL_iXlinker.Device_2_EtherCAT.Term_9_EK1100.Term_10_EK1122.Term_18_EK1100.Term_22_EL3011.AI_Standard.Status/TxPDO_Toggle <-> AI Standard/Status/TxPDO Toggle
//     PlcTask Inputs/GVL_iXlinker.Device_2_EtherCAT.Term_9_EK1100.Term_10_EK1122.Term_18_EK1100.Term_22_EL3011.AI_Standard.Status/Underrange <-> AI Standard/Status/Underrange
//     PlcTask Inputs/GVL_iXlinker.Device_2_EtherCAT.Term_9_EK1100.Term_10_EK1122.Term_18_EK1100.Term_22_EL3011.AI_Standard.Value <-> AI Standard/Value
//     PlcTask Inputs/GVL_iXlinker.Device_2_EtherCAT.Term_9_EK1100.Term_10_EK1122.Term_18_EK1100.Term_22_EL3011.InfoData.AdsAddr <-> InfoData/AdsAddr
//     PlcTask Inputs/GVL_iXlinker.Device_2_EtherCAT.Term_9_EK1100.Term_10_EK1122.Term_18_EK1100.Term_22_EL3011.InfoData.State <-> InfoData/State
//     PlcTask Inputs/GVL_iXlinker.Device_2_EtherCAT.Term_9_EK1100.Term_10_EK1122.Term_18_EK1100.Term_22_EL3011.WcState.InputToggle <-> WcState/InputToggle
//     PlcTask Inputs/GVL_iXlinker.Device_2_EtherCAT.Term_9_EK1100.Term_10_EK1122.Term_18_EK1100.Term_22_EL3011.WcState.WcState <-> WcState/WcState
//   TcoIoTests/TcoIoTests Instance <-> Device 2 (EtherCAT)/Term 9 (EK1100)/Term 10 (EK1122)/Term 23 (EK1100)
//     PlcTask Inputs/GVL_iXlinker.Device_2_EtherCAT.Term_9_EK1100.Term_10_EK1122.Term_23_EK1100.InfoData.State <-> InfoData/State
//   TcoIoTests/TcoIoTests Instance <-> Device 2 (EtherCAT)/Term 9 (EK1100)/Term 10 (EK1122)/Term 23 (EK1100)/Term 24 (EK1122)
//     PlcTask Inputs/GVL_iXlinker.Device_2_EtherCAT.Term_9_EK1100.Term_10_EK1122.Term_23_EK1100.Term_24_EK1122.InfoData.State <-> InfoData/State
//   TcoIoTests/TcoIoTests Instance <-> Device 2 (EtherCAT)/Term 9 (EK1100)/Term 10 (EK1122)/Term 23 (EK1100)/Term 24 (EK1122)/Term 25 (EK1100)
//     PlcTask Inputs/GVL_iXlinker.Device_2_EtherCAT.Term_9_EK1100.Term_10_EK1122.Term_23_EK1100.Term_24_EK1122.Term_25_EK1100.InfoData.State <-> InfoData/State
//   TcoIoTests/TcoIoTests Instance <-> Device 2 (EtherCAT)/Term 9 (EK1100)/Term 10 (EK1122)/Term 23 (EK1100)/Term 24 (EK1122)/Term 25 (EK1100)/Term 26 (EL1819)
//     PlcTask Inputs/GVL_iXlinker.Device_2_EtherCAT.Term_9_EK1100.Term_10_EK1122.Term_23_EK1100.Term_24_EK1122.Term_25_EK1100.Term_26_EL1819.Channel_{1..16}.Input <-> Channel {1..16}/Input  (16 links)
//     PlcTask Inputs/GVL_iXlinker.Device_2_EtherCAT.Term_9_EK1100.Term_10_EK1122.Term_23_EK1100.Term_24_EK1122.Term_25_EK1100.Term_26_EL1819.InfoData.State <-> InfoData/State
//     PlcTask Inputs/GVL_iXlinker.Device_2_EtherCAT.Term_9_EK1100.Term_10_EK1122.Term_23_EK1100.Term_24_EK1122.Term_25_EK1100.Term_26_EL1819.WcState.InputToggle <-> WcState/InputToggle
//     PlcTask Inputs/GVL_iXlinker.Device_2_EtherCAT.Term_9_EK1100.Term_10_EK1122.Term_23_EK1100.Term_24_EK1122.Term_25_EK1100.Term_26_EL1819.WcState.WcState <-> WcState/WcState
//   TcoIoTests/TcoIoTests Instance <-> Device 2 (EtherCAT)/Term 9 (EK1100)/Term 10 (EK1122)/Term 23 (EK1100)/Term 24 (EK1122)/Term 25 (EK1100)/Term 27 (EL1819)
//     PlcTask Inputs/GVL_iXlinker.Device_2_EtherCAT.Term_9_EK1100.Term_10_EK1122.Term_23_EK1100.Term_24_EK1122.Term_25_EK1100.Term_27_EL1819.Channel_{1..16}.Input <-> Channel {1..16}/Input  (16 links)
//     PlcTask Inputs/GVL_iXlinker.Device_2_EtherCAT.Term_9_EK1100.Term_10_EK1122.Term_23_EK1100.Term_24_EK1122.Term_25_EK1100.Term_27_EL1819.InfoData.State <-> InfoData/State
//     PlcTask Inputs/GVL_iXlinker.Device_2_EtherCAT.Term_9_EK1100.Term_10_EK1122.Term_23_EK1100.Term_24_EK1122.Term_25_EK1100.Term_27_EL1819.WcState.InputToggle <-> WcState/InputToggle
//     PlcTask Inputs/GVL_iXlinker.Device_2_EtherCAT.Term_9_EK1100.Term_10_EK1122.Term_23_EK1100.Term_24_EK1122.Term_25_EK1100.Term_27_EL1819.WcState.WcState <-> WcState/WcState
//   TcoIoTests/TcoIoTests Instance <-> Device 2 (EtherCAT)/Term 9 (EK1100)/Term 10 (EK1122)/Term 23 (EK1100)/Term 24 (EK1122)/Term 28 (EK1100)
//     PlcTask Inputs/GVL_iXlinker.Device_2_EtherCAT.Term_9_EK1100.Term_10_EK1122.Term_23_EK1100.Term_24_EK1122.Term_28_EK1100.InfoData.State <-> InfoData/State
//   TcoIoTests/TcoIoTests Instance <-> Device 2 (EtherCAT)/Term 9 (EK1100)/Term 10 (EK1122)/Term 23 (EK1100)/Term 24 (EK1122)/Term 28 (EK1100)/Term 29 (EL2788)
//     PlcTask Inputs/GVL_iXlinker.Device_2_EtherCAT.Term_9_EK1100.Term_10_EK1122.Term_23_EK1100.Term_24_EK1122.Term_28_EK1100.Term_29_EL2788.InfoData.State <-> InfoData/State
//     PlcTask Inputs/GVL_iXlinker.Device_2_EtherCAT.Term_9_EK1100.Term_10_EK1122.Term_23_EK1100.Term_24_EK1122.Term_28_EK1100.Term_29_EL2788.WcState.WcState <-> WcState/WcState
//     PlcTask Outputs/GVL_iXlinker.Device_2_EtherCAT.Term_9_EK1100.Term_10_EK1122.Term_23_EK1100.Term_24_EK1122.Term_28_EK1100.Term_29_EL2788.Channel_{1..8}.Output <-> Channel {1..8}/Output  (8 links)
//   TcoIoTests/TcoIoTests Instance <-> Device 2 (EtherCAT)/Term 9 (EK1100)/Term 10 (EK1122)/Term 23 (EK1100)/Term 24 (EK1122)/Term 28 (EK1100)/Term 30 (EL3773)
//     PlcTask Inputs/GVL_iXlinker.Device_2_EtherCAT.Term_9_EK1100.Term_10_EK1122.Term_23_EK1100.Term_24_EK1122.Term_28_EK1100.Term_30_EL3773.AI_NextSync1Time.StartTimeNextLatch/Hi <-> AI NextSync1Time/StartTimeNextLatch/Hi
//     PlcTask Inputs/GVL_iXlinker.Device_2_EtherCAT.Term_9_EK1100.Term_10_EK1122.Term_23_EK1100.Term_24_EK1122.Term_28_EK1100.Term_30_EL3773.AI_NextSync1Time.StartTimeNextLatch/Low <-> AI NextSync1Time/StartTimeNextLatch/Low
//     PlcTask Inputs/GVL_iXlinker.Device_2_EtherCAT.Term_9_EK1100.Term_10_EK1122.Term_23_EK1100.Term_24_EK1122.Term_28_EK1100.Term_30_EL3773.AI_Sample_Count.Sample_Count <-> AI Sample Count/Sample Count
//     PlcTask Inputs/GVL_iXlinker.Device_2_EtherCAT.Term_9_EK1100.Term_10_EK1122.Term_23_EK1100.Term_24_EK1122.Term_28_EK1100.Term_30_EL3773.InfoData.AdsAddr <-> InfoData/AdsAddr
//     PlcTask Inputs/GVL_iXlinker.Device_2_EtherCAT.Term_9_EK1100.Term_10_EK1122.Term_23_EK1100.Term_24_EK1122.Term_28_EK1100.Term_30_EL3773.InfoData.DcInputShift <-> InfoData/DcInputShift
//     PlcTask Inputs/GVL_iXlinker.Device_2_EtherCAT.Term_9_EK1100.Term_10_EK1122.Term_23_EK1100.Term_24_EK1122.Term_28_EK1100.Term_30_EL3773.InfoData.DcOutputShift <-> InfoData/DcOutputShift
//     PlcTask Inputs/GVL_iXlinker.Device_2_EtherCAT.Term_9_EK1100.Term_10_EK1122.Term_23_EK1100.Term_24_EK1122.Term_28_EK1100.Term_30_EL3773.InfoData.State <-> InfoData/State
//     PlcTask Inputs/GVL_iXlinker.Device_2_EtherCAT.Term_9_EK1100.Term_10_EK1122.Term_23_EK1100.Term_24_EK1122.Term_28_EK1100.Term_30_EL3773.L1_Current_Status.I1_Status/Error <-> L1 Current Status/I1 Status/Error
//     PlcTask Inputs/GVL_iXlinker.Device_2_EtherCAT.Term_9_EK1100.Term_10_EK1122.Term_23_EK1100.Term_24_EK1122.Term_28_EK1100.Term_30_EL3773.L2_Current_Status.I2_Status/Error <-> L2 Current Status/I2 Status/Error
//     PlcTask Inputs/GVL_iXlinker.Device_2_EtherCAT.Term_9_EK1100.Term_10_EK1122.Term_23_EK1100.Term_24_EK1122.Term_28_EK1100.Term_30_EL3773.L3_Current_Status.I3_Status/Error <-> L3 Current Status/I3 Status/Error
//     PlcTask Inputs/GVL_iXlinker.Device_2_EtherCAT.Term_9_EK1100.Term_10_EK1122.Term_23_EK1100.Term_24_EK1122.Term_28_EK1100.Term_30_EL3773.L1_Current_Status.I1_Status/Limit_x <-> L1 Current Status/I1 Status/Limit
//     PlcTask Inputs/GVL_iXlinker.Device_2_EtherCAT.Term_9_EK1100.Term_10_EK1122.Term_23_EK1100.Term_24_EK1122.Term_28_EK1100.Term_30_EL3773.L2_Current_Status.I2_Status/Limit_x <-> L2 Current Status/I2 Status/Limit
//     PlcTask Inputs/GVL_iXlinker.Device_2_EtherCAT.Term_9_EK1100.Term_10_EK1122.Term_23_EK1100.Term_24_EK1122.Term_28_EK1100.Term_30_EL3773.L3_Current_Status.I3_Status/Limit_x <-> L3 Current Status/I3 Status/Limit
//     PlcTask Inputs/GVL_iXlinker.Device_2_EtherCAT.Term_9_EK1100.Term_10_EK1122.Term_23_EK1100.Term_24_EK1122.Term_28_EK1100.Term_30_EL3773.L1_Current_Status.I1_Status/Overrange <-> L1 Current Status/I1 Status/Overrange
//     PlcTask Inputs/GVL_iXlinker.Device_2_EtherCAT.Term_9_EK1100.Term_10_EK1122.Term_23_EK1100.Term_24_EK1122.Term_28_EK1100.Term_30_EL3773.L2_Current_Status.I2_Status/Overrange <-> L2 Current Status/I2 Status/Overrange
//     PlcTask Inputs/GVL_iXlinker.Device_2_EtherCAT.Term_9_EK1100.Term_10_EK1122.Term_23_EK1100.Term_24_EK1122.Term_28_EK1100.Term_30_EL3773.L3_Current_Status.I3_Status/Overrange <-> L3 Current Status/I3 Status/Overrange
//     PlcTask Inputs/GVL_iXlinker.Device_2_EtherCAT.Term_9_EK1100.Term_10_EK1122.Term_23_EK1100.Term_24_EK1122.Term_28_EK1100.Term_30_EL3773.L1_Current_Status.I1_Status/Sync_error <-> L1 Current Status/I1 Status/Sync error
//     PlcTask Inputs/GVL_iXlinker.Device_2_EtherCAT.Term_9_EK1100.Term_10_EK1122.Term_23_EK1100.Term_24_EK1122.Term_28_EK1100.Term_30_EL3773.L2_Current_Status.I2_Status/Sync_error <-> L2 Current Status/I2 Status/Sync error
//     PlcTask Inputs/GVL_iXlinker.Device_2_EtherCAT.Term_9_EK1100.Term_10_EK1122.Term_23_EK1100.Term_24_EK1122.Term_28_EK1100.Term_30_EL3773.L3_Current_Status.I3_Status/Sync_error <-> L3 Current Status/I3 Status/Sync error
//     PlcTask Inputs/GVL_iXlinker.Device_2_EtherCAT.Term_9_EK1100.Term_10_EK1122.Term_23_EK1100.Term_24_EK1122.Term_28_EK1100.Term_30_EL3773.L1_Current_Status.I1_Status/TxPDO_State <-> L1 Current Status/I1 Status/TxPDO State
//     PlcTask Inputs/GVL_iXlinker.Device_2_EtherCAT.Term_9_EK1100.Term_10_EK1122.Term_23_EK1100.Term_24_EK1122.Term_28_EK1100.Term_30_EL3773.L2_Current_Status.I2_Status/TxPDO_State <-> L2 Current Status/I2 Status/TxPDO State
//     PlcTask Inputs/GVL_iXlinker.Device_2_EtherCAT.Term_9_EK1100.Term_10_EK1122.Term_23_EK1100.Term_24_EK1122.Term_28_EK1100.Term_30_EL3773.L3_Current_Status.I3_Status/TxPDO_State <-> L3 Current Status/I3 Status/TxPDO State
//     PlcTask Inputs/GVL_iXlinker.Device_2_EtherCAT.Term_9_EK1100.Term_10_EK1122.Term_23_EK1100.Term_24_EK1122.Term_28_EK1100.Term_30_EL3773.L1_Current_Status.I1_Status/TxPDO_Toggle <-> L1 Current Status/I1 Status/TxPDO Toggle
//     PlcTask Inputs/GVL_iXlinker.Device_2_EtherCAT.Term_9_EK1100.Term_10_EK1122.Term_23_EK1100.Term_24_EK1122.Term_28_EK1100.Term_30_EL3773.L2_Current_Status.I2_Status/TxPDO_Toggle <-> L2 Current Status/I2 Status/TxPDO Toggle
//     PlcTask Inputs/GVL_iXlinker.Device_2_EtherCAT.Term_9_EK1100.Term_10_EK1122.Term_23_EK1100.Term_24_EK1122.Term_28_EK1100.Term_30_EL3773.L3_Current_Status.I3_Status/TxPDO_Toggle <-> L3 Current Status/I3 Status/TxPDO Toggle
//     PlcTask Inputs/GVL_iXlinker.Device_2_EtherCAT.Term_9_EK1100.Term_10_EK1122.Term_23_EK1100.Term_24_EK1122.Term_28_EK1100.Term_30_EL3773.L1_Current_Status.I1_Status/Underrange <-> L1 Current Status/I1 Status/Underrange
//     PlcTask Inputs/GVL_iXlinker.Device_2_EtherCAT.Term_9_EK1100.Term_10_EK1122.Term_23_EK1100.Term_24_EK1122.Term_28_EK1100.Term_30_EL3773.L2_Current_Status.I2_Status/Underrange <-> L2 Current Status/I2 Status/Underrange
//     PlcTask Inputs/GVL_iXlinker.Device_2_EtherCAT.Term_9_EK1100.Term_10_EK1122.Term_23_EK1100.Term_24_EK1122.Term_28_EK1100.Term_30_EL3773.L3_Current_Status.I3_Status/Underrange <-> L3 Current Status/I3 Status/Underrange
//     PlcTask Inputs/GVL_iXlinker.Device_2_EtherCAT.Term_9_EK1100.Term_10_EK1122.Term_23_EK1100.Term_24_EK1122.Term_28_EK1100.Term_30_EL3773.L1_Voltage_Status.U1_Status/Error <-> L1 Voltage Status/U1 Status/Error
//     PlcTask Inputs/GVL_iXlinker.Device_2_EtherCAT.Term_9_EK1100.Term_10_EK1122.Term_23_EK1100.Term_24_EK1122.Term_28_EK1100.Term_30_EL3773.L2_Voltage_Status.U2_Status/Error <-> L2 Voltage Status/U2 Status/Error
//     PlcTask Inputs/GVL_iXlinker.Device_2_EtherCAT.Term_9_EK1100.Term_10_EK1122.Term_23_EK1100.Term_24_EK1122.Term_28_EK1100.Term_30_EL3773.L3_Voltage_Status.U3_Status/Error <-> L3 Voltage Status/U3 Status/Error
//     PlcTask Inputs/GVL_iXlinker.Device_2_EtherCAT.Term_9_EK1100.Term_10_EK1122.Term_23_EK1100.Term_24_EK1122.Term_28_EK1100.Term_30_EL3773.L1_Voltage_Status.U1_Status/Limit_x <-> L1 Voltage Status/U1 Status/Limit
//     PlcTask Inputs/GVL_iXlinker.Device_2_EtherCAT.Term_9_EK1100.Term_10_EK1122.Term_23_EK1100.Term_24_EK1122.Term_28_EK1100.Term_30_EL3773.L2_Voltage_Status.U2_Status/Limit_x <-> L2 Voltage Status/U2 Status/Limit
//     PlcTask Inputs/GVL_iXlinker.Device_2_EtherCAT.Term_9_EK1100.Term_10_EK1122.Term_23_EK1100.Term_24_EK1122.Term_28_EK1100.Term_30_EL3773.L3_Voltage_Status.U3_Status/Limit_x <-> L3 Voltage Status/U3 Status/Limit
//     PlcTask Inputs/GVL_iXlinker.Device_2_EtherCAT.Term_9_EK1100.Term_10_EK1122.Term_23_EK1100.Term_24_EK1122.Term_28_EK1100.Term_30_EL3773.L1_Voltage_Status.U1_Status/Overrange <-> L1 Voltage Status/U1 Status/Overrange
//     PlcTask Inputs/GVL_iXlinker.Device_2_EtherCAT.Term_9_EK1100.Term_10_EK1122.Term_23_EK1100.Term_24_EK1122.Term_28_EK1100.Term_30_EL3773.L2_Voltage_Status.U2_Status/Overrange <-> L2 Voltage Status/U2 Status/Overrange
//     PlcTask Inputs/GVL_iXlinker.Device_2_EtherCAT.Term_9_EK1100.Term_10_EK1122.Term_23_EK1100.Term_24_EK1122.Term_28_EK1100.Term_30_EL3773.L3_Voltage_Status.U3_Status/Overrange <-> L3 Voltage Status/U3 Status/Overrange
//     PlcTask Inputs/GVL_iXlinker.Device_2_EtherCAT.Term_9_EK1100.Term_10_EK1122.Term_23_EK1100.Term_24_EK1122.Term_28_EK1100.Term_30_EL3773.L1_Voltage_Status.U1_Status/Sync_error <-> L1 Voltage Status/U1 Status/Sync error
//     PlcTask Inputs/GVL_iXlinker.Device_2_EtherCAT.Term_9_EK1100.Term_10_EK1122.Term_23_EK1100.Term_24_EK1122.Term_28_EK1100.Term_30_EL3773.L2_Voltage_Status.U2_Status/Sync_error <-> L2 Voltage Status/U2 Status/Sync error
//     PlcTask Inputs/GVL_iXlinker.Device_2_EtherCAT.Term_9_EK1100.Term_10_EK1122.Term_23_EK1100.Term_24_EK1122.Term_28_EK1100.Term_30_EL3773.L3_Voltage_Status.U3_Status/Sync_error <-> L3 Voltage Status/U3 Status/Sync error
//     PlcTask Inputs/GVL_iXlinker.Device_2_EtherCAT.Term_9_EK1100.Term_10_EK1122.Term_23_EK1100.Term_24_EK1122.Term_28_EK1100.Term_30_EL3773.L1_Voltage_Status.U1_Status/TxPDO_State <-> L1 Voltage Status/U1 Status/TxPDO State
//     PlcTask Inputs/GVL_iXlinker.Device_2_EtherCAT.Term_9_EK1100.Term_10_EK1122.Term_23_EK1100.Term_24_EK1122.Term_28_EK1100.Term_30_EL3773.L2_Voltage_Status.U2_Status/TxPDO_State <-> L2 Voltage Status/U2 Status/TxPDO State
//     PlcTask Inputs/GVL_iXlinker.Device_2_EtherCAT.Term_9_EK1100.Term_10_EK1122.Term_23_EK1100.Term_24_EK1122.Term_28_EK1100.Term_30_EL3773.L3_Voltage_Status.U3_Status/TxPDO_State <-> L3 Voltage Status/U3 Status/TxPDO State
//     PlcTask Inputs/GVL_iXlinker.Device_2_EtherCAT.Term_9_EK1100.Term_10_EK1122.Term_23_EK1100.Term_24_EK1122.Term_28_EK1100.Term_30_EL3773.L1_Voltage_Status.U1_Status/TxPDO_Toggle <-> L1 Voltage Status/U1 Status/TxPDO Toggle
//     PlcTask Inputs/GVL_iXlinker.Device_2_EtherCAT.Term_9_EK1100.Term_10_EK1122.Term_23_EK1100.Term_24_EK1122.Term_28_EK1100.Term_30_EL3773.L2_Voltage_Status.U2_Status/TxPDO_Toggle <-> L2 Voltage Status/U2 Status/TxPDO Toggle
//     PlcTask Inputs/GVL_iXlinker.Device_2_EtherCAT.Term_9_EK1100.Term_10_EK1122.Term_23_EK1100.Term_24_EK1122.Term_28_EK1100.Term_30_EL3773.L3_Voltage_Status.U3_Status/TxPDO_Toggle <-> L3 Voltage Status/U3 Status/TxPDO Toggle
//     PlcTask Inputs/GVL_iXlinker.Device_2_EtherCAT.Term_9_EK1100.Term_10_EK1122.Term_23_EK1100.Term_24_EK1122.Term_28_EK1100.Term_30_EL3773.L1_Voltage_Status.U1_Status/Underrange <-> L1 Voltage Status/U1 Status/Underrange
//     PlcTask Inputs/GVL_iXlinker.Device_2_EtherCAT.Term_9_EK1100.Term_10_EK1122.Term_23_EK1100.Term_24_EK1122.Term_28_EK1100.Term_30_EL3773.L2_Voltage_Status.U2_Status/Underrange <-> L2 Voltage Status/U2 Status/Underrange
//     PlcTask Inputs/GVL_iXlinker.Device_2_EtherCAT.Term_9_EK1100.Term_10_EK1122.Term_23_EK1100.Term_24_EK1122.Term_28_EK1100.Term_30_EL3773.L3_Voltage_Status.U3_Status/Underrange <-> L3 Voltage Status/U3 Status/Underrange
//     PlcTask Inputs/GVL_iXlinker.Device_2_EtherCAT.Term_9_EK1100.Term_10_EK1122.Term_23_EK1100.Term_24_EK1122.Term_28_EK1100.Term_30_EL3773.WcState.InputToggle <-> WcState/InputToggle
//     PlcTask Inputs/GVL_iXlinker.Device_2_EtherCAT.Term_9_EK1100.Term_10_EK1122.Term_23_EK1100.Term_24_EK1122.Term_28_EK1100.Term_30_EL3773.WcState.WcState <-> WcState/WcState
//   TcoIoTests/TcoIoTests Instance <-> Device 2 (EtherCAT)/Term 9 (EK1100)/Term 10 (EK1122)/Term 23 (EK1100)/Term 31 (EL3773)
//     PlcTask Inputs/GVL_iXlinker.Device_2_EtherCAT.Term_9_EK1100.Term_10_EK1122.Term_23_EK1100.Term_31_EL3773.AI_NextSync1Time.StartTimeNextLatch/Hi <-> AI NextSync1Time/StartTimeNextLatch/Hi
//     PlcTask Inputs/GVL_iXlinker.Device_2_EtherCAT.Term_9_EK1100.Term_10_EK1122.Term_23_EK1100.Term_31_EL3773.AI_NextSync1Time.StartTimeNextLatch/Low <-> AI NextSync1Time/StartTimeNextLatch/Low
//     PlcTask Inputs/GVL_iXlinker.Device_2_EtherCAT.Term_9_EK1100.Term_10_EK1122.Term_23_EK1100.Term_31_EL3773.AI_Sample_Count.Sample_Count <-> AI Sample Count/Sample Count
//     PlcTask Inputs/GVL_iXlinker.Device_2_EtherCAT.Term_9_EK1100.Term_10_EK1122.Term_23_EK1100.Term_31_EL3773.InfoData.AdsAddr <-> InfoData/AdsAddr
//     PlcTask Inputs/GVL_iXlinker.Device_2_EtherCAT.Term_9_EK1100.Term_10_EK1122.Term_23_EK1100.Term_31_EL3773.InfoData.DcInputShift <-> InfoData/DcInputShift
//     PlcTask Inputs/GVL_iXlinker.Device_2_EtherCAT.Term_9_EK1100.Term_10_EK1122.Term_23_EK1100.Term_31_EL3773.InfoData.DcOutputShift <-> InfoData/DcOutputShift
//     PlcTask Inputs/GVL_iXlinker.Device_2_EtherCAT.Term_9_EK1100.Term_10_EK1122.Term_23_EK1100.Term_31_EL3773.InfoData.State <-> InfoData/State
//     PlcTask Inputs/GVL_iXlinker.Device_2_EtherCAT.Term_9_EK1100.Term_10_EK1122.Term_23_EK1100.Term_31_EL3773.L1_Current_Status.I1_Status/Error <-> L1 Current Status/I1 Status/Error
//     PlcTask Inputs/GVL_iXlinker.Device_2_EtherCAT.Term_9_EK1100.Term_10_EK1122.Term_23_EK1100.Term_31_EL3773.L2_Current_Status.I2_Status/Error <-> L2 Current Status/I2 Status/Error
//     PlcTask Inputs/GVL_iXlinker.Device_2_EtherCAT.Term_9_EK1100.Term_10_EK1122.Term_23_EK1100.Term_31_EL3773.L3_Current_Status.I3_Status/Error <-> L3 Current Status/I3 Status/Error
//     PlcTask Inputs/GVL_iXlinker.Device_2_EtherCAT.Term_9_EK1100.Term_10_EK1122.Term_23_EK1100.Term_31_EL3773.L1_Current_Status.I1_Status/Limit_x <-> L1 Current Status/I1 Status/Limit
//     PlcTask Inputs/GVL_iXlinker.Device_2_EtherCAT.Term_9_EK1100.Term_10_EK1122.Term_23_EK1100.Term_31_EL3773.L2_Current_Status.I2_Status/Limit_x <-> L2 Current Status/I2 Status/Limit
//     PlcTask Inputs/GVL_iXlinker.Device_2_EtherCAT.Term_9_EK1100.Term_10_EK1122.Term_23_EK1100.Term_31_EL3773.L3_Current_Status.I3_Status/Limit_x <-> L3 Current Status/I3 Status/Limit
//     PlcTask Inputs/GVL_iXlinker.Device_2_EtherCAT.Term_9_EK1100.Term_10_EK1122.Term_23_EK1100.Term_31_EL3773.L1_Current_Status.I1_Status/Overrange <-> L1 Current Status/I1 Status/Overrange
//     PlcTask Inputs/GVL_iXlinker.Device_2_EtherCAT.Term_9_EK1100.Term_10_EK1122.Term_23_EK1100.Term_31_EL3773.L2_Current_Status.I2_Status/Overrange <-> L2 Current Status/I2 Status/Overrange
//     PlcTask Inputs/GVL_iXlinker.Device_2_EtherCAT.Term_9_EK1100.Term_10_EK1122.Term_23_EK1100.Term_31_EL3773.L3_Current_Status.I3_Status/Overrange <-> L3 Current Status/I3 Status/Overrange
//     PlcTask Inputs/GVL_iXlinker.Device_2_EtherCAT.Term_9_EK1100.Term_10_EK1122.Term_23_EK1100.Term_31_EL3773.L1_Current_Status.I1_Status/Sync_error <-> L1 Current Status/I1 Status/Sync error
//     PlcTask Inputs/GVL_iXlinker.Device_2_EtherCAT.Term_9_EK1100.Term_10_EK1122.Term_23_EK1100.Term_31_EL3773.L2_Current_Status.I2_Status/Sync_error <-> L2 Current Status/I2 Status/Sync error
//     PlcTask Inputs/GVL_iXlinker.Device_2_EtherCAT.Term_9_EK1100.Term_10_EK1122.Term_23_EK1100.Term_31_EL3773.L3_Current_Status.I3_Status/Sync_error <-> L3 Current Status/I3 Status/Sync error
//     PlcTask Inputs/GVL_iXlinker.Device_2_EtherCAT.Term_9_EK1100.Term_10_EK1122.Term_23_EK1100.Term_31_EL3773.L1_Current_Status.I1_Status/TxPDO_State <-> L1 Current Status/I1 Status/TxPDO State
//     PlcTask Inputs/GVL_iXlinker.Device_2_EtherCAT.Term_9_EK1100.Term_10_EK1122.Term_23_EK1100.Term_31_EL3773.L2_Current_Status.I2_Status/TxPDO_State <-> L2 Current Status/I2 Status/TxPDO State
//     PlcTask Inputs/GVL_iXlinker.Device_2_EtherCAT.Term_9_EK1100.Term_10_EK1122.Term_23_EK1100.Term_31_EL3773.L3_Current_Status.I3_Status/TxPDO_State <-> L3 Current Status/I3 Status/TxPDO State
//     PlcTask Inputs/GVL_iXlinker.Device_2_EtherCAT.Term_9_EK1100.Term_10_EK1122.Term_23_EK1100.Term_31_EL3773.L1_Current_Status.I1_Status/TxPDO_Toggle <-> L1 Current Status/I1 Status/TxPDO Toggle
//     PlcTask Inputs/GVL_iXlinker.Device_2_EtherCAT.Term_9_EK1100.Term_10_EK1122.Term_23_EK1100.Term_31_EL3773.L2_Current_Status.I2_Status/TxPDO_Toggle <-> L2 Current Status/I2 Status/TxPDO Toggle
//     PlcTask Inputs/GVL_iXlinker.Device_2_EtherCAT.Term_9_EK1100.Term_10_EK1122.Term_23_EK1100.Term_31_EL3773.L3_Current_Status.I3_Status/TxPDO_Toggle <-> L3 Current Status/I3 Status/TxPDO Toggle
//     PlcTask Inputs/GVL_iXlinker.Device_2_EtherCAT.Term_9_EK1100.Term_10_EK1122.Term_23_EK1100.Term_31_EL3773.L1_Current_Status.I1_Status/Underrange <-> L1 Current Status/I1 Status/Underrange
//     PlcTask Inputs/GVL_iXlinker.Device_2_EtherCAT.Term_9_EK1100.Term_10_EK1122.Term_23_EK1100.Term_31_EL3773.L2_Current_Status.I2_Status/Underrange <-> L2 Current Status/I2 Status/Underrange
//     PlcTask Inputs/GVL_iXlinker.Device_2_EtherCAT.Term_9_EK1100.Term_10_EK1122.Term_23_EK1100.Term_31_EL3773.L3_Current_Status.I3_Status/Underrange <-> L3 Current Status/I3 Status/Underrange
//     PlcTask Inputs/GVL_iXlinker.Device_2_EtherCAT.Term_9_EK1100.Term_10_EK1122.Term_23_EK1100.Term_31_EL3773.L1_Voltage_Status.U1_Status/Error <-> L1 Voltage Status/U1 Status/Error
//     PlcTask Inputs/GVL_iXlinker.Device_2_EtherCAT.Term_9_EK1100.Term_10_EK1122.Term_23_EK1100.Term_31_EL3773.L2_Voltage_Status.U2_Status/Error <-> L2 Voltage Status/U2 Status/Error
//     PlcTask Inputs/GVL_iXlinker.Device_2_EtherCAT.Term_9_EK1100.Term_10_EK1122.Term_23_EK1100.Term_31_EL3773.L3_Voltage_Status.U3_Status/Error <-> L3 Voltage Status/U3 Status/Error
//     PlcTask Inputs/GVL_iXlinker.Device_2_EtherCAT.Term_9_EK1100.Term_10_EK1122.Term_23_EK1100.Term_31_EL3773.L1_Voltage_Status.U1_Status/Limit_x <-> L1 Voltage Status/U1 Status/Limit
//     PlcTask Inputs/GVL_iXlinker.Device_2_EtherCAT.Term_9_EK1100.Term_10_EK1122.Term_23_EK1100.Term_31_EL3773.L2_Voltage_Status.U2_Status/Limit_x <-> L2 Voltage Status/U2 Status/Limit
//     PlcTask Inputs/GVL_iXlinker.Device_2_EtherCAT.Term_9_EK1100.Term_10_EK1122.Term_23_EK1100.Term_31_EL3773.L3_Voltage_Status.U3_Status/Limit_x <-> L3 Voltage Status/U3 Status/Limit
//     PlcTask Inputs/GVL_iXlinker.Device_2_EtherCAT.Term_9_EK1100.Term_10_EK1122.Term_23_EK1100.Term_31_EL3773.L1_Voltage_Status.U1_Status/Overrange <-> L1 Voltage Status/U1 Status/Overrange
//     PlcTask Inputs/GVL_iXlinker.Device_2_EtherCAT.Term_9_EK1100.Term_10_EK1122.Term_23_EK1100.Term_31_EL3773.L2_Voltage_Status.U2_Status/Overrange <-> L2 Voltage Status/U2 Status/Overrange
//     PlcTask Inputs/GVL_iXlinker.Device_2_EtherCAT.Term_9_EK1100.Term_10_EK1122.Term_23_EK1100.Term_31_EL3773.L3_Voltage_Status.U3_Status/Overrange <-> L3 Voltage Status/U3 Status/Overrange
//     PlcTask Inputs/GVL_iXlinker.Device_2_EtherCAT.Term_9_EK1100.Term_10_EK1122.Term_23_EK1100.Term_31_EL3773.L1_Voltage_Status.U1_Status/Sync_error <-> L1 Voltage Status/U1 Status/Sync error
//     PlcTask Inputs/GVL_iXlinker.Device_2_EtherCAT.Term_9_EK1100.Term_10_EK1122.Term_23_EK1100.Term_31_EL3773.L2_Voltage_Status.U2_Status/Sync_error <-> L2 Voltage Status/U2 Status/Sync error
//     PlcTask Inputs/GVL_iXlinker.Device_2_EtherCAT.Term_9_EK1100.Term_10_EK1122.Term_23_EK1100.Term_31_EL3773.L3_Voltage_Status.U3_Status/Sync_error <-> L3 Voltage Status/U3 Status/Sync error
//     PlcTask Inputs/GVL_iXlinker.Device_2_EtherCAT.Term_9_EK1100.Term_10_EK1122.Term_23_EK1100.Term_31_EL3773.L1_Voltage_Status.U1_Status/TxPDO_State <-> L1 Voltage Status/U1 Status/TxPDO State
//     PlcTask Inputs/GVL_iXlinker.Device_2_EtherCAT.Term_9_EK1100.Term_10_EK1122.Term_23_EK1100.Term_31_EL3773.L2_Voltage_Status.U2_Status/TxPDO_State <-> L2 Voltage Status/U2 Status/TxPDO State
//     PlcTask Inputs/GVL_iXlinker.Device_2_EtherCAT.Term_9_EK1100.Term_10_EK1122.Term_23_EK1100.Term_31_EL3773.L3_Voltage_Status.U3_Status/TxPDO_State <-> L3 Voltage Status/U3 Status/TxPDO State
//     PlcTask Inputs/GVL_iXlinker.Device_2_EtherCAT.Term_9_EK1100.Term_10_EK1122.Term_23_EK1100.Term_31_EL3773.L1_Voltage_Status.U1_Status/TxPDO_Toggle <-> L1 Voltage Status/U1 Status/TxPDO Toggle
//     PlcTask Inputs/GVL_iXlinker.Device_2_EtherCAT.Term_9_EK1100.Term_10_EK1122.Term_23_EK1100.Term_31_EL3773.L2_Voltage_Status.U2_Status/TxPDO_Toggle <-> L2 Voltage Status/U2 Status/TxPDO Toggle
//     PlcTask Inputs/GVL_iXlinker.Device_2_EtherCAT.Term_9_EK1100.Term_10_EK1122.Term_23_EK1100.Term_31_EL3773.L3_Voltage_Status.U3_Status/TxPDO_Toggle <-> L3 Voltage Status/U3 Status/TxPDO Toggle
//     PlcTask Inputs/GVL_iXlinker.Device_2_EtherCAT.Term_9_EK1100.Term_10_EK1122.Term_23_EK1100.Term_31_EL3773.L1_Voltage_Status.U1_Status/Underrange <-> L1 Voltage Status/U1 Status/Underrange
//     PlcTask Inputs/GVL_iXlinker.Device_2_EtherCAT.Term_9_EK1100.Term_10_EK1122.Term_23_EK1100.Term_31_EL3773.L2_Voltage_Status.U2_Status/Underrange <-> L2 Voltage Status/U2 Status/Underrange
//     PlcTask Inputs/GVL_iXlinker.Device_2_EtherCAT.Term_9_EK1100.Term_10_EK1122.Term_23_EK1100.Term_31_EL3773.L3_Voltage_Status.U3_Status/Underrange <-> L3 Voltage Status/U3 Status/Underrange
//     PlcTask Inputs/GVL_iXlinker.Device_2_EtherCAT.Term_9_EK1100.Term_10_EK1122.Term_23_EK1100.Term_31_EL3773.WcState.InputToggle <-> WcState/InputToggle
//     PlcTask Inputs/GVL_iXlinker.Device_2_EtherCAT.Term_9_EK1100.Term_10_EK1122.Term_23_EK1100.Term_31_EL3773.WcState.WcState <-> WcState/WcState
//   TcoIoTests/TcoIoTests Instance <-> Device 2 (EtherCAT)/Term 9 (EK1100)/Term 10 (EK1122)/Term 23 (EK1100)/Term 32 (EL2258)
//     PlcTask Inputs/GVL_iXlinker.Device_2_EtherCAT.Term_9_EK1100.Term_10_EK1122.Term_23_EK1100.Term_32_EL2258.InfoData.AdsAddr <-> InfoData/AdsAddr
//     PlcTask Inputs/GVL_iXlinker.Device_2_EtherCAT.Term_9_EK1100.Term_10_EK1122.Term_23_EK1100.Term_32_EL2258.InfoData.DcInputShift <-> InfoData/DcInputShift
//     PlcTask Inputs/GVL_iXlinker.Device_2_EtherCAT.Term_9_EK1100.Term_10_EK1122.Term_23_EK1100.Term_32_EL2258.InfoData.DcOutputShift <-> InfoData/DcOutputShift
//     PlcTask Inputs/GVL_iXlinker.Device_2_EtherCAT.Term_9_EK1100.Term_10_EK1122.Term_23_EK1100.Term_32_EL2258.InfoData.State <-> InfoData/State
//     PlcTask Inputs/GVL_iXlinker.Device_2_EtherCAT.Term_9_EK1100.Term_10_EK1122.Term_23_EK1100.Term_32_EL2258.MTO_Inputs_Channel_{1..8}.Status/Events_in_output_buffer <-> MTO Inputs Channel {1..8}/Status/Events in output buffer  (8 links)
//     PlcTask Inputs/GVL_iXlinker.Device_2_EtherCAT.Term_9_EK1100.Term_10_EK1122.Term_23_EK1100.Term_32_EL2258.MTO_Inputs_Channel_{1..8}.Status/Input_cycle_counter <-> MTO Inputs Channel {1..8}/Status/Input cycle counter  (8 links)
//     PlcTask Inputs/GVL_iXlinker.Device_2_EtherCAT.Term_9_EK1100.Term_10_EK1122.Term_23_EK1100.Term_32_EL2258.MTO_Inputs_Channel_{1..8}.Status/Output_buffer_overflow <-> MTO Inputs Channel {1..8}/Status/Output buffer overflow  (8 links)
//     PlcTask Inputs/GVL_iXlinker.Device_2_EtherCAT.Term_9_EK1100.Term_10_EK1122.Term_23_EK1100.Term_32_EL2258.MTO_Inputs_Channel_{1..8}.Status/Output_order_feedback <-> MTO Inputs Channel {1..8}/Status/Output order feedback  (8 links)
//     PlcTask Inputs/GVL_iXlinker.Device_2_EtherCAT.Term_9_EK1100.Term_10_EK1122.Term_23_EK1100.Term_32_EL2258.MTO_Inputs_Channel_{1..8}.Status/Output_short_circuit <-> MTO Inputs Channel {1..8}/Status/Output short circuit  (8 links)
//     PlcTask Inputs/GVL_iXlinker.Device_2_EtherCAT.Term_9_EK1100.Term_10_EK1122.Term_23_EK1100.Term_32_EL2258.MTO_Inputs_Channel_{1..8}.Status/Output_state <-> MTO Inputs Channel {1..8}/Status/Output state  (8 links)
//     PlcTask Inputs/GVL_iXlinker.Device_2_EtherCAT.Term_9_EK1100.Term_10_EK1122.Term_23_EK1100.Term_32_EL2258.WcState.InputToggle <-> WcState/InputToggle
//     PlcTask Inputs/GVL_iXlinker.Device_2_EtherCAT.Term_9_EK1100.Term_10_EK1122.Term_23_EK1100.Term_32_EL2258.WcState.WcState <-> WcState/WcState
//     PlcTask Outputs/GVL_iXlinker.Device_2_EtherCAT.Term_9_EK1100.Term_10_EK1122.Term_23_EK1100.Term_32_EL2258.MTO_Outputs_10x_Channel_{1..8}.Ctrl/Enable_manual_operation <-> MTO Outputs 10x Channel {1..8}/Ctrl/Enable manual operation  (8 links)
//     PlcTask Outputs/GVL_iXlinker.Device_2_EtherCAT.Term_9_EK1100.Term_10_EK1122.Term_23_EK1100.Term_32_EL2258.MTO_Outputs_10x_Channel_{1..8}.Ctrl/Force_order <-> MTO Outputs 10x Channel {1..8}/Ctrl/Force order  (8 links)
//     PlcTask Outputs/GVL_iXlinker.Device_2_EtherCAT.Term_9_EK1100.Term_10_EK1122.Term_23_EK1100.Term_32_EL2258.MTO_Outputs_10x_Channel_{1..8}.Ctrl/Manual_output_state <-> MTO Outputs 10x Channel {1..8}/Ctrl/Manual output state  (8 links)
//     PlcTask Outputs/GVL_iXlinker.Device_2_EtherCAT.Term_9_EK1100.Term_10_EK1122.Term_23_EK1100.Term_32_EL2258.MTO_Outputs_10x_Channel_{1..8}.Ctrl/No_of_output_events <-> MTO Outputs 10x Channel {1..8}/Ctrl/No of output events  (8 links)
//     PlcTask Outputs/GVL_iXlinker.Device_2_EtherCAT.Term_9_EK1100.Term_10_EK1122.Term_23_EK1100.Term_32_EL2258.MTO_Outputs_10x_Channel_{1..8}.Ctrl/Output_buffer_reset <-> MTO Outputs 10x Channel {1..8}/Ctrl/Output buffer reset  (8 links)
//     PlcTask Outputs/GVL_iXlinker.Device_2_EtherCAT.Term_9_EK1100.Term_10_EK1122.Term_23_EK1100.Term_32_EL2258.MTO_Outputs_10x_Channel_{1..8}.Ctrl/Output_order_counter <-> MTO Outputs 10x Channel {1..8}/Ctrl/Output order counter  (8 links)
//     PlcTask Outputs/GVL_iXlinker.Device_2_EtherCAT.Term_9_EK1100.Term_10_EK1122.Term_23_EK1100.Term_32_EL2258.MTO_Outputs_10x_Channel_1.Output_event_time[0] <-> MTO Outputs 10x Channel 1/Output event time 1
//     PlcTask Outputs/GVL_iXlinker.Device_2_EtherCAT.Term_9_EK1100.Term_10_EK1122.Term_23_EK1100.Term_32_EL2258.MTO_Outputs_10x_Channel_1.Output_event_time[1] <-> MTO Outputs 10x Channel 1/Output event time 2
//     PlcTask Outputs/GVL_iXlinker.Device_2_EtherCAT.Term_9_EK1100.Term_10_EK1122.Term_23_EK1100.Term_32_EL2258.MTO_Outputs_10x_Channel_1.Output_event_time[2] <-> MTO Outputs 10x Channel 1/Output event time 3
//     PlcTask Outputs/GVL_iXlinker.Device_2_EtherCAT.Term_9_EK1100.Term_10_EK1122.Term_23_EK1100.Term_32_EL2258.MTO_Outputs_10x_Channel_1.Output_event_time[3] <-> MTO Outputs 10x Channel 1/Output event time 4
//     PlcTask Outputs/GVL_iXlinker.Device_2_EtherCAT.Term_9_EK1100.Term_10_EK1122.Term_23_EK1100.Term_32_EL2258.MTO_Outputs_10x_Channel_1.Output_event_time[4] <-> MTO Outputs 10x Channel 1/Output event time 5
//     PlcTask Outputs/GVL_iXlinker.Device_2_EtherCAT.Term_9_EK1100.Term_10_EK1122.Term_23_EK1100.Term_32_EL2258.MTO_Outputs_10x_Channel_1.Output_event_time[5] <-> MTO Outputs 10x Channel 1/Output event time 6
//     PlcTask Outputs/GVL_iXlinker.Device_2_EtherCAT.Term_9_EK1100.Term_10_EK1122.Term_23_EK1100.Term_32_EL2258.MTO_Outputs_10x_Channel_1.Output_event_time[6] <-> MTO Outputs 10x Channel 1/Output event time 7
//     PlcTask Outputs/GVL_iXlinker.Device_2_EtherCAT.Term_9_EK1100.Term_10_EK1122.Term_23_EK1100.Term_32_EL2258.MTO_Outputs_10x_Channel_1.Output_event_time[7] <-> MTO Outputs 10x Channel 1/Output event time 8
//     PlcTask Outputs/GVL_iXlinker.Device_2_EtherCAT.Term_9_EK1100.Term_10_EK1122.Term_23_EK1100.Term_32_EL2258.MTO_Outputs_10x_Channel_1.Output_event_time[8] <-> MTO Outputs 10x Channel 1/Output event time 9
//     PlcTask Outputs/GVL_iXlinker.Device_2_EtherCAT.Term_9_EK1100.Term_10_EK1122.Term_23_EK1100.Term_32_EL2258.MTO_Outputs_10x_Channel_1.Output_event_time[9] <-> MTO Outputs 10x Channel 1/Output event time 10
//     PlcTask Outputs/GVL_iXlinker.Device_2_EtherCAT.Term_9_EK1100.Term_10_EK1122.Term_23_EK1100.Term_32_EL2258.MTO_Outputs_10x_Channel_2.Output_event_time[0] <-> MTO Outputs 10x Channel 2/Output event time 1
//     PlcTask Outputs/GVL_iXlinker.Device_2_EtherCAT.Term_9_EK1100.Term_10_EK1122.Term_23_EK1100.Term_32_EL2258.MTO_Outputs_10x_Channel_2.Output_event_time[1] <-> MTO Outputs 10x Channel 2/Output event time 2
//     PlcTask Outputs/GVL_iXlinker.Device_2_EtherCAT.Term_9_EK1100.Term_10_EK1122.Term_23_EK1100.Term_32_EL2258.MTO_Outputs_10x_Channel_2.Output_event_time[2] <-> MTO Outputs 10x Channel 2/Output event time 3
//     PlcTask Outputs/GVL_iXlinker.Device_2_EtherCAT.Term_9_EK1100.Term_10_EK1122.Term_23_EK1100.Term_32_EL2258.MTO_Outputs_10x_Channel_2.Output_event_time[3] <-> MTO Outputs 10x Channel 2/Output event time 4
//     PlcTask Outputs/GVL_iXlinker.Device_2_EtherCAT.Term_9_EK1100.Term_10_EK1122.Term_23_EK1100.Term_32_EL2258.MTO_Outputs_10x_Channel_2.Output_event_time[4] <-> MTO Outputs 10x Channel 2/Output event time 5
//     PlcTask Outputs/GVL_iXlinker.Device_2_EtherCAT.Term_9_EK1100.Term_10_EK1122.Term_23_EK1100.Term_32_EL2258.MTO_Outputs_10x_Channel_2.Output_event_time[5] <-> MTO Outputs 10x Channel 2/Output event time 6
//     PlcTask Outputs/GVL_iXlinker.Device_2_EtherCAT.Term_9_EK1100.Term_10_EK1122.Term_23_EK1100.Term_32_EL2258.MTO_Outputs_10x_Channel_2.Output_event_time[6] <-> MTO Outputs 10x Channel 2/Output event time 7
//     PlcTask Outputs/GVL_iXlinker.Device_2_EtherCAT.Term_9_EK1100.Term_10_EK1122.Term_23_EK1100.Term_32_EL2258.MTO_Outputs_10x_Channel_2.Output_event_time[7] <-> MTO Outputs 10x Channel 2/Output event time 8
//     PlcTask Outputs/GVL_iXlinker.Device_2_EtherCAT.Term_9_EK1100.Term_10_EK1122.Term_23_EK1100.Term_32_EL2258.MTO_Outputs_10x_Channel_2.Output_event_time[8] <-> MTO Outputs 10x Channel 2/Output event time 9
//     PlcTask Outputs/GVL_iXlinker.Device_2_EtherCAT.Term_9_EK1100.Term_10_EK1122.Term_23_EK1100.Term_32_EL2258.MTO_Outputs_10x_Channel_2.Output_event_time[9] <-> MTO Outputs 10x Channel 2/Output event time 10
//     PlcTask Outputs/GVL_iXlinker.Device_2_EtherCAT.Term_9_EK1100.Term_10_EK1122.Term_23_EK1100.Term_32_EL2258.MTO_Outputs_10x_Channel_3.Output_event_time[0] <-> MTO Outputs 10x Channel 3/Output event time 1
//     PlcTask Outputs/GVL_iXlinker.Device_2_EtherCAT.Term_9_EK1100.Term_10_EK1122.Term_23_EK1100.Term_32_EL2258.MTO_Outputs_10x_Channel_3.Output_event_time[1] <-> MTO Outputs 10x Channel 3/Output event time 2
//     PlcTask Outputs/GVL_iXlinker.Device_2_EtherCAT.Term_9_EK1100.Term_10_EK1122.Term_23_EK1100.Term_32_EL2258.MTO_Outputs_10x_Channel_3.Output_event_time[2] <-> MTO Outputs 10x Channel 3/Output event time 3
//     PlcTask Outputs/GVL_iXlinker.Device_2_EtherCAT.Term_9_EK1100.Term_10_EK1122.Term_23_EK1100.Term_32_EL2258.MTO_Outputs_10x_Channel_3.Output_event_time[3] <-> MTO Outputs 10x Channel 3/Output event time 4
//     PlcTask Outputs/GVL_iXlinker.Device_2_EtherCAT.Term_9_EK1100.Term_10_EK1122.Term_23_EK1100.Term_32_EL2258.MTO_Outputs_10x_Channel_3.Output_event_time[4] <-> MTO Outputs 10x Channel 3/Output event time 5
//     PlcTask Outputs/GVL_iXlinker.Device_2_EtherCAT.Term_9_EK1100.Term_10_EK1122.Term_23_EK1100.Term_32_EL2258.MTO_Outputs_10x_Channel_3.Output_event_time[5] <-> MTO Outputs 10x Channel 3/Output event time 6
//     PlcTask Outputs/GVL_iXlinker.Device_2_EtherCAT.Term_9_EK1100.Term_10_EK1122.Term_23_EK1100.Term_32_EL2258.MTO_Outputs_10x_Channel_3.Output_event_time[6] <-> MTO Outputs 10x Channel 3/Output event time 7
//     PlcTask Outputs/GVL_iXlinker.Device_2_EtherCAT.Term_9_EK1100.Term_10_EK1122.Term_23_EK1100.Term_32_EL2258.MTO_Outputs_10x_Channel_3.Output_event_time[7] <-> MTO Outputs 10x Channel 3/Output event time 8
//     PlcTask Outputs/GVL_iXlinker.Device_2_EtherCAT.Term_9_EK1100.Term_10_EK1122.Term_23_EK1100.Term_32_EL2258.MTO_Outputs_10x_Channel_3.Output_event_time[8] <-> MTO Outputs 10x Channel 3/Output event time 9
//     PlcTask Outputs/GVL_iXlinker.Device_2_EtherCAT.Term_9_EK1100.Term_10_EK1122.Term_23_EK1100.Term_32_EL2258.MTO_Outputs_10x_Channel_3.Output_event_time[9] <-> MTO Outputs 10x Channel 3/Output event time 10
//     PlcTask Outputs/GVL_iXlinker.Device_2_EtherCAT.Term_9_EK1100.Term_10_EK1122.Term_23_EK1100.Term_32_EL2258.MTO_Outputs_10x_Channel_4.Output_event_time[0] <-> MTO Outputs 10x Channel 4/Output event time 1
//     PlcTask Outputs/GVL_iXlinker.Device_2_EtherCAT.Term_9_EK1100.Term_10_EK1122.Term_23_EK1100.Term_32_EL2258.MTO_Outputs_10x_Channel_4.Output_event_time[1] <-> MTO Outputs 10x Channel 4/Output event time 2
//     PlcTask Outputs/GVL_iXlinker.Device_2_EtherCAT.Term_9_EK1100.Term_10_EK1122.Term_23_EK1100.Term_32_EL2258.MTO_Outputs_10x_Channel_4.Output_event_time[2] <-> MTO Outputs 10x Channel 4/Output event time 3
//     PlcTask Outputs/GVL_iXlinker.Device_2_EtherCAT.Term_9_EK1100.Term_10_EK1122.Term_23_EK1100.Term_32_EL2258.MTO_Outputs_10x_Channel_4.Output_event_time[3] <-> MTO Outputs 10x Channel 4/Output event time 4
//     PlcTask Outputs/GVL_iXlinker.Device_2_EtherCAT.Term_9_EK1100.Term_10_EK1122.Term_23_EK1100.Term_32_EL2258.MTO_Outputs_10x_Channel_4.Output_event_time[4] <-> MTO Outputs 10x Channel 4/Output event time 5
//     PlcTask Outputs/GVL_iXlinker.Device_2_EtherCAT.Term_9_EK1100.Term_10_EK1122.Term_23_EK1100.Term_32_EL2258.MTO_Outputs_10x_Channel_4.Output_event_time[5] <-> MTO Outputs 10x Channel 4/Output event time 6
//     PlcTask Outputs/GVL_iXlinker.Device_2_EtherCAT.Term_9_EK1100.Term_10_EK1122.Term_23_EK1100.Term_32_EL2258.MTO_Outputs_10x_Channel_4.Output_event_time[6] <-> MTO Outputs 10x Channel 4/Output event time 7
//     PlcTask Outputs/GVL_iXlinker.Device_2_EtherCAT.Term_9_EK1100.Term_10_EK1122.Term_23_EK1100.Term_32_EL2258.MTO_Outputs_10x_Channel_4.Output_event_time[7] <-> MTO Outputs 10x Channel 4/Output event time 8
//     PlcTask Outputs/GVL_iXlinker.Device_2_EtherCAT.Term_9_EK1100.Term_10_EK1122.Term_23_EK1100.Term_32_EL2258.MTO_Outputs_10x_Channel_4.Output_event_time[8] <-> MTO Outputs 10x Channel 4/Output event time 9
//     PlcTask Outputs/GVL_iXlinker.Device_2_EtherCAT.Term_9_EK1100.Term_10_EK1122.Term_23_EK1100.Term_32_EL2258.MTO_Outputs_10x_Channel_4.Output_event_time[9] <-> MTO Outputs 10x Channel 4/Output event time 10
//     PlcTask Outputs/GVL_iXlinker.Device_2_EtherCAT.Term_9_EK1100.Term_10_EK1122.Term_23_EK1100.Term_32_EL2258.MTO_Outputs_10x_Channel_5.Output_event_time[0] <-> MTO Outputs 10x Channel 5/Output event time 1
//     PlcTask Outputs/GVL_iXlinker.Device_2_EtherCAT.Term_9_EK1100.Term_10_EK1122.Term_23_EK1100.Term_32_EL2258.MTO_Outputs_10x_Channel_5.Output_event_time[1] <-> MTO Outputs 10x Channel 5/Output event time 2
//     PlcTask Outputs/GVL_iXlinker.Device_2_EtherCAT.Term_9_EK1100.Term_10_EK1122.Term_23_EK1100.Term_32_EL2258.MTO_Outputs_10x_Channel_5.Output_event_time[2] <-> MTO Outputs 10x Channel 5/Output event time 3
//     PlcTask Outputs/GVL_iXlinker.Device_2_EtherCAT.Term_9_EK1100.Term_10_EK1122.Term_23_EK1100.Term_32_EL2258.MTO_Outputs_10x_Channel_5.Output_event_time[3] <-> MTO Outputs 10x Channel 5/Output event time 4
//     PlcTask Outputs/GVL_iXlinker.Device_2_EtherCAT.Term_9_EK1100.Term_10_EK1122.Term_23_EK1100.Term_32_EL2258.MTO_Outputs_10x_Channel_5.Output_event_time[4] <-> MTO Outputs 10x Channel 5/Output event time 5
//     PlcTask Outputs/GVL_iXlinker.Device_2_EtherCAT.Term_9_EK1100.Term_10_EK1122.Term_23_EK1100.Term_32_EL2258.MTO_Outputs_10x_Channel_5.Output_event_time[5] <-> MTO Outputs 10x Channel 5/Output event time 6
//     PlcTask Outputs/GVL_iXlinker.Device_2_EtherCAT.Term_9_EK1100.Term_10_EK1122.Term_23_EK1100.Term_32_EL2258.MTO_Outputs_10x_Channel_5.Output_event_time[6] <-> MTO Outputs 10x Channel 5/Output event time 7
//     PlcTask Outputs/GVL_iXlinker.Device_2_EtherCAT.Term_9_EK1100.Term_10_EK1122.Term_23_EK1100.Term_32_EL2258.MTO_Outputs_10x_Channel_5.Output_event_time[7] <-> MTO Outputs 10x Channel 5/Output event time 8
//     PlcTask Outputs/GVL_iXlinker.Device_2_EtherCAT.Term_9_EK1100.Term_10_EK1122.Term_23_EK1100.Term_32_EL2258.MTO_Outputs_10x_Channel_5.Output_event_time[8] <-> MTO Outputs 10x Channel 5/Output event time 9
//     PlcTask Outputs/GVL_iXlinker.Device_2_EtherCAT.Term_9_EK1100.Term_10_EK1122.Term_23_EK1100.Term_32_EL2258.MTO_Outputs_10x_Channel_5.Output_event_time[9] <-> MTO Outputs 10x Channel 5/Output event time 10
//     PlcTask Outputs/GVL_iXlinker.Device_2_EtherCAT.Term_9_EK1100.Term_10_EK1122.Term_23_EK1100.Term_32_EL2258.MTO_Outputs_10x_Channel_6.Output_event_time[0] <-> MTO Outputs 10x Channel 6/Output event time 1
//     PlcTask Outputs/GVL_iXlinker.Device_2_EtherCAT.Term_9_EK1100.Term_10_EK1122.Term_23_EK1100.Term_32_EL2258.MTO_Outputs_10x_Channel_6.Output_event_time[1] <-> MTO Outputs 10x Channel 6/Output event time 2
//     PlcTask Outputs/GVL_iXlinker.Device_2_EtherCAT.Term_9_EK1100.Term_10_EK1122.Term_23_EK1100.Term_32_EL2258.MTO_Outputs_10x_Channel_6.Output_event_time[2] <-> MTO Outputs 10x Channel 6/Output event time 3
//     PlcTask Outputs/GVL_iXlinker.Device_2_EtherCAT.Term_9_EK1100.Term_10_EK1122.Term_23_EK1100.Term_32_EL2258.MTO_Outputs_10x_Channel_6.Output_event_time[3] <-> MTO Outputs 10x Channel 6/Output event time 4
//     PlcTask Outputs/GVL_iXlinker.Device_2_EtherCAT.Term_9_EK1100.Term_10_EK1122.Term_23_EK1100.Term_32_EL2258.MTO_Outputs_10x_Channel_6.Output_event_time[4] <-> MTO Outputs 10x Channel 6/Output event time 5
//     PlcTask Outputs/GVL_iXlinker.Device_2_EtherCAT.Term_9_EK1100.Term_10_EK1122.Term_23_EK1100.Term_32_EL2258.MTO_Outputs_10x_Channel_6.Output_event_time[5] <-> MTO Outputs 10x Channel 6/Output event time 6
//     PlcTask Outputs/GVL_iXlinker.Device_2_EtherCAT.Term_9_EK1100.Term_10_EK1122.Term_23_EK1100.Term_32_EL2258.MTO_Outputs_10x_Channel_6.Output_event_time[6] <-> MTO Outputs 10x Channel 6/Output event time 7
//     PlcTask Outputs/GVL_iXlinker.Device_2_EtherCAT.Term_9_EK1100.Term_10_EK1122.Term_23_EK1100.Term_32_EL2258.MTO_Outputs_10x_Channel_6.Output_event_time[7] <-> MTO Outputs 10x Channel 6/Output event time 8
//     PlcTask Outputs/GVL_iXlinker.Device_2_EtherCAT.Term_9_EK1100.Term_10_EK1122.Term_23_EK1100.Term_32_EL2258.MTO_Outputs_10x_Channel_6.Output_event_time[8] <-> MTO Outputs 10x Channel 6/Output event time 9
//     PlcTask Outputs/GVL_iXlinker.Device_2_EtherCAT.Term_9_EK1100.Term_10_EK1122.Term_23_EK1100.Term_32_EL2258.MTO_Outputs_10x_Channel_6.Output_event_time[9] <-> MTO Outputs 10x Channel 6/Output event time 10
//     PlcTask Outputs/GVL_iXlinker.Device_2_EtherCAT.Term_9_EK1100.Term_10_EK1122.Term_23_EK1100.Term_32_EL2258.MTO_Outputs_10x_Channel_7.Output_event_time[0] <-> MTO Outputs 10x Channel 7/Output event time 1
//     PlcTask Outputs/GVL_iXlinker.Device_2_EtherCAT.Term_9_EK1100.Term_10_EK1122.Term_23_EK1100.Term_32_EL2258.MTO_Outputs_10x_Channel_7.Output_event_time[1] <-> MTO Outputs 10x Channel 7/Output event time 2
//     PlcTask Outputs/GVL_iXlinker.Device_2_EtherCAT.Term_9_EK1100.Term_10_EK1122.Term_23_EK1100.Term_32_EL2258.MTO_Outputs_10x_Channel_7.Output_event_time[2] <-> MTO Outputs 10x Channel 7/Output event time 3
//     PlcTask Outputs/GVL_iXlinker.Device_2_EtherCAT.Term_9_EK1100.Term_10_EK1122.Term_23_EK1100.Term_32_EL2258.MTO_Outputs_10x_Channel_7.Output_event_time[3] <-> MTO Outputs 10x Channel 7/Output event time 4
//     PlcTask Outputs/GVL_iXlinker.Device_2_EtherCAT.Term_9_EK1100.Term_10_EK1122.Term_23_EK1100.Term_32_EL2258.MTO_Outputs_10x_Channel_7.Output_event_time[4] <-> MTO Outputs 10x Channel 7/Output event time 5
//     PlcTask Outputs/GVL_iXlinker.Device_2_EtherCAT.Term_9_EK1100.Term_10_EK1122.Term_23_EK1100.Term_32_EL2258.MTO_Outputs_10x_Channel_7.Output_event_time[5] <-> MTO Outputs 10x Channel 7/Output event time 6
//     PlcTask Outputs/GVL_iXlinker.Device_2_EtherCAT.Term_9_EK1100.Term_10_EK1122.Term_23_EK1100.Term_32_EL2258.MTO_Outputs_10x_Channel_7.Output_event_time[6] <-> MTO Outputs 10x Channel 7/Output event time 7
//     PlcTask Outputs/GVL_iXlinker.Device_2_EtherCAT.Term_9_EK1100.Term_10_EK1122.Term_23_EK1100.Term_32_EL2258.MTO_Outputs_10x_Channel_7.Output_event_time[7] <-> MTO Outputs 10x Channel 7/Output event time 8
//     PlcTask Outputs/GVL_iXlinker.Device_2_EtherCAT.Term_9_EK1100.Term_10_EK1122.Term_23_EK1100.Term_32_EL2258.MTO_Outputs_10x_Channel_7.Output_event_time[8] <-> MTO Outputs 10x Channel 7/Output event time 9
//     PlcTask Outputs/GVL_iXlinker.Device_2_EtherCAT.Term_9_EK1100.Term_10_EK1122.Term_23_EK1100.Term_32_EL2258.MTO_Outputs_10x_Channel_7.Output_event_time[9] <-> MTO Outputs 10x Channel 7/Output event time 10
//     PlcTask Outputs/GVL_iXlinker.Device_2_EtherCAT.Term_9_EK1100.Term_10_EK1122.Term_23_EK1100.Term_32_EL2258.MTO_Outputs_10x_Channel_8.Output_event_time[0] <-> MTO Outputs 10x Channel 8/Output event time 1
//     PlcTask Outputs/GVL_iXlinker.Device_2_EtherCAT.Term_9_EK1100.Term_10_EK1122.Term_23_EK1100.Term_32_EL2258.MTO_Outputs_10x_Channel_8.Output_event_time[1] <-> MTO Outputs 10x Channel 8/Output event time 2
//     PlcTask Outputs/GVL_iXlinker.Device_2_EtherCAT.Term_9_EK1100.Term_10_EK1122.Term_23_EK1100.Term_32_EL2258.MTO_Outputs_10x_Channel_8.Output_event_time[2] <-> MTO Outputs 10x Channel 8/Output event time 3
//     PlcTask Outputs/GVL_iXlinker.Device_2_EtherCAT.Term_9_EK1100.Term_10_EK1122.Term_23_EK1100.Term_32_EL2258.MTO_Outputs_10x_Channel_8.Output_event_time[3] <-> MTO Outputs 10x Channel 8/Output event time 4
//     PlcTask Outputs/GVL_iXlinker.Device_2_EtherCAT.Term_9_EK1100.Term_10_EK1122.Term_23_EK1100.Term_32_EL2258.MTO_Outputs_10x_Channel_8.Output_event_time[4] <-> MTO Outputs 10x Channel 8/Output event time 5
//     PlcTask Outputs/GVL_iXlinker.Device_2_EtherCAT.Term_9_EK1100.Term_10_EK1122.Term_23_EK1100.Term_32_EL2258.MTO_Outputs_10x_Channel_8.Output_event_time[5] <-> MTO Outputs 10x Channel 8/Output event time 6
//     PlcTask Outputs/GVL_iXlinker.Device_2_EtherCAT.Term_9_EK1100.Term_10_EK1122.Term_23_EK1100.Term_32_EL2258.MTO_Outputs_10x_Channel_8.Output_event_time[6] <-> MTO Outputs 10x Channel 8/Output event time 7
//     PlcTask Outputs/GVL_iXlinker.Device_2_EtherCAT.Term_9_EK1100.Term_10_EK1122.Term_23_EK1100.Term_32_EL2258.MTO_Outputs_10x_Channel_8.Output_event_time[7] <-> MTO Outputs 10x Channel 8/Output event time 8
//     PlcTask Outputs/GVL_iXlinker.Device_2_EtherCAT.Term_9_EK1100.Term_10_EK1122.Term_23_EK1100.Term_32_EL2258.MTO_Outputs_10x_Channel_8.Output_event_time[8] <-> MTO Outputs 10x Channel 8/Output event time 9
//     PlcTask Outputs/GVL_iXlinker.Device_2_EtherCAT.Term_9_EK1100.Term_10_EK1122.Term_23_EK1100.Term_32_EL2258.MTO_Outputs_10x_Channel_8.Output_event_time[9] <-> MTO Outputs 10x Channel 8/Output event time 10
//     PlcTask Outputs/GVL_iXlinker.Device_2_EtherCAT.Term_9_EK1100.Term_10_EK1122.Term_23_EK1100.Term_32_EL2258.MTO_Outputs_10x_Channel_1.Outputs/Output_event_state_1 <-> MTO Outputs 10x Channel 1/Outputs/Output event state 1
//     PlcTask Outputs/GVL_iXlinker.Device_2_EtherCAT.Term_9_EK1100.Term_10_EK1122.Term_23_EK1100.Term_32_EL2258.MTO_Outputs_10x_Channel_1.Outputs/Output_event_state_10 <-> MTO Outputs 10x Channel 1/Outputs/Output event state 10
//     PlcTask Outputs/GVL_iXlinker.Device_2_EtherCAT.Term_9_EK1100.Term_10_EK1122.Term_23_EK1100.Term_32_EL2258.MTO_Outputs_10x_Channel_1.Outputs/Output_event_state_2 <-> MTO Outputs 10x Channel 1/Outputs/Output event state 2
//     PlcTask Outputs/GVL_iXlinker.Device_2_EtherCAT.Term_9_EK1100.Term_10_EK1122.Term_23_EK1100.Term_32_EL2258.MTO_Outputs_10x_Channel_1.Outputs/Output_event_state_3 <-> MTO Outputs 10x Channel 1/Outputs/Output event state 3
//     PlcTask Outputs/GVL_iXlinker.Device_2_EtherCAT.Term_9_EK1100.Term_10_EK1122.Term_23_EK1100.Term_32_EL2258.MTO_Outputs_10x_Channel_1.Outputs/Output_event_state_4 <-> MTO Outputs 10x Channel 1/Outputs/Output event state 4
//     PlcTask Outputs/GVL_iXlinker.Device_2_EtherCAT.Term_9_EK1100.Term_10_EK1122.Term_23_EK1100.Term_32_EL2258.MTO_Outputs_10x_Channel_1.Outputs/Output_event_state_5 <-> MTO Outputs 10x Channel 1/Outputs/Output event state 5
//     PlcTask Outputs/GVL_iXlinker.Device_2_EtherCAT.Term_9_EK1100.Term_10_EK1122.Term_23_EK1100.Term_32_EL2258.MTO_Outputs_10x_Channel_1.Outputs/Output_event_state_6 <-> MTO Outputs 10x Channel 1/Outputs/Output event state 6
//     PlcTask Outputs/GVL_iXlinker.Device_2_EtherCAT.Term_9_EK1100.Term_10_EK1122.Term_23_EK1100.Term_32_EL2258.MTO_Outputs_10x_Channel_1.Outputs/Output_event_state_7 <-> MTO Outputs 10x Channel 1/Outputs/Output event state 7
//     PlcTask Outputs/GVL_iXlinker.Device_2_EtherCAT.Term_9_EK1100.Term_10_EK1122.Term_23_EK1100.Term_32_EL2258.MTO_Outputs_10x_Channel_1.Outputs/Output_event_state_8 <-> MTO Outputs 10x Channel 1/Outputs/Output event state 8
//     PlcTask Outputs/GVL_iXlinker.Device_2_EtherCAT.Term_9_EK1100.Term_10_EK1122.Term_23_EK1100.Term_32_EL2258.MTO_Outputs_10x_Channel_1.Outputs/Output_event_state_9 <-> MTO Outputs 10x Channel 1/Outputs/Output event state 9
//     PlcTask Outputs/GVL_iXlinker.Device_2_EtherCAT.Term_9_EK1100.Term_10_EK1122.Term_23_EK1100.Term_32_EL2258.MTO_Outputs_10x_Channel_2.Outputs/Output_event_state_1 <-> MTO Outputs 10x Channel 2/Outputs/Output event state 1
//     PlcTask Outputs/GVL_iXlinker.Device_2_EtherCAT.Term_9_EK1100.Term_10_EK1122.Term_23_EK1100.Term_32_EL2258.MTO_Outputs_10x_Channel_2.Outputs/Output_event_state_10 <-> MTO Outputs 10x Channel 2/Outputs/Output event state 10
//     PlcTask Outputs/GVL_iXlinker.Device_2_EtherCAT.Term_9_EK1100.Term_10_EK1122.Term_23_EK1100.Term_32_EL2258.MTO_Outputs_10x_Channel_2.Outputs/Output_event_state_2 <-> MTO Outputs 10x Channel 2/Outputs/Output event state 2
//     PlcTask Outputs/GVL_iXlinker.Device_2_EtherCAT.Term_9_EK1100.Term_10_EK1122.Term_23_EK1100.Term_32_EL2258.MTO_Outputs_10x_Channel_2.Outputs/Output_event_state_3 <-> MTO Outputs 10x Channel 2/Outputs/Output event state 3
//     PlcTask Outputs/GVL_iXlinker.Device_2_EtherCAT.Term_9_EK1100.Term_10_EK1122.Term_23_EK1100.Term_32_EL2258.MTO_Outputs_10x_Channel_2.Outputs/Output_event_state_4 <-> MTO Outputs 10x Channel 2/Outputs/Output event state 4
//     PlcTask Outputs/GVL_iXlinker.Device_2_EtherCAT.Term_9_EK1100.Term_10_EK1122.Term_23_EK1100.Term_32_EL2258.MTO_Outputs_10x_Channel_2.Outputs/Output_event_state_5 <-> MTO Outputs 10x Channel 2/Outputs/Output event state 5
//     PlcTask Outputs/GVL_iXlinker.Device_2_EtherCAT.Term_9_EK1100.Term_10_EK1122.Term_23_EK1100.Term_32_EL2258.MTO_Outputs_10x_Channel_2.Outputs/Output_event_state_6 <-> MTO Outputs 10x Channel 2/Outputs/Output event state 6
//     PlcTask Outputs/GVL_iXlinker.Device_2_EtherCAT.Term_9_EK1100.Term_10_EK1122.Term_23_EK1100.Term_32_EL2258.MTO_Outputs_10x_Channel_2.Outputs/Output_event_state_7 <-> MTO Outputs 10x Channel 2/Outputs/Output event state 7
//     PlcTask Outputs/GVL_iXlinker.Device_2_EtherCAT.Term_9_EK1100.Term_10_EK1122.Term_23_EK1100.Term_32_EL2258.MTO_Outputs_10x_Channel_2.Outputs/Output_event_state_8 <-> MTO Outputs 10x Channel 2/Outputs/Output event state 8
//     PlcTask Outputs/GVL_iXlinker.Device_2_EtherCAT.Term_9_EK1100.Term_10_EK1122.Term_23_EK1100.Term_32_EL2258.MTO_Outputs_10x_Channel_2.Outputs/Output_event_state_9 <-> MTO Outputs 10x Channel 2/Outputs/Output event state 9
//     PlcTask Outputs/GVL_iXlinker.Device_2_EtherCAT.Term_9_EK1100.Term_10_EK1122.Term_23_EK1100.Term_32_EL2258.MTO_Outputs_10x_Channel_3.Outputs/Output_event_state_1 <-> MTO Outputs 10x Channel 3/Outputs/Output event state 1
//     PlcTask Outputs/GVL_iXlinker.Device_2_EtherCAT.Term_9_EK1100.Term_10_EK1122.Term_23_EK1100.Term_32_EL2258.MTO_Outputs_10x_Channel_3.Outputs/Output_event_state_10 <-> MTO Outputs 10x Channel 3/Outputs/Output event state 10
//     PlcTask Outputs/GVL_iXlinker.Device_2_EtherCAT.Term_9_EK1100.Term_10_EK1122.Term_23_EK1100.Term_32_EL2258.MTO_Outputs_10x_Channel_3.Outputs/Output_event_state_2 <-> MTO Outputs 10x Channel 3/Outputs/Output event state 2
//     PlcTask Outputs/GVL_iXlinker.Device_2_EtherCAT.Term_9_EK1100.Term_10_EK1122.Term_23_EK1100.Term_32_EL2258.MTO_Outputs_10x_Channel_3.Outputs/Output_event_state_3 <-> MTO Outputs 10x Channel 3/Outputs/Output event state 3
//     PlcTask Outputs/GVL_iXlinker.Device_2_EtherCAT.Term_9_EK1100.Term_10_EK1122.Term_23_EK1100.Term_32_EL2258.MTO_Outputs_10x_Channel_3.Outputs/Output_event_state_4 <-> MTO Outputs 10x Channel 3/Outputs/Output event state 4
//     PlcTask Outputs/GVL_iXlinker.Device_2_EtherCAT.Term_9_EK1100.Term_10_EK1122.Term_23_EK1100.Term_32_EL2258.MTO_Outputs_10x_Channel_3.Outputs/Output_event_state_5 <-> MTO Outputs 10x Channel 3/Outputs/Output event state 5
//     PlcTask Outputs/GVL_iXlinker.Device_2_EtherCAT.Term_9_EK1100.Term_10_EK1122.Term_23_EK1100.Term_32_EL2258.MTO_Outputs_10x_Channel_3.Outputs/Output_event_state_6 <-> MTO Outputs 10x Channel 3/Outputs/Output event state 6
//     PlcTask Outputs/GVL_iXlinker.Device_2_EtherCAT.Term_9_EK1100.Term_10_EK1122.Term_23_EK1100.Term_32_EL2258.MTO_Outputs_10x_Channel_3.Outputs/Output_event_state_7 <-> MTO Outputs 10x Channel 3/Outputs/Output event state 7
//     PlcTask Outputs/GVL_iXlinker.Device_2_EtherCAT.Term_9_EK1100.Term_10_EK1122.Term_23_EK1100.Term_32_EL2258.MTO_Outputs_10x_Channel_3.Outputs/Output_event_state_8 <-> MTO Outputs 10x Channel 3/Outputs/Output event state 8
//     PlcTask Outputs/GVL_iXlinker.Device_2_EtherCAT.Term_9_EK1100.Term_10_EK1122.Term_23_EK1100.Term_32_EL2258.MTO_Outputs_10x_Channel_3.Outputs/Output_event_state_9 <-> MTO Outputs 10x Channel 3/Outputs/Output event state 9
//     PlcTask Outputs/GVL_iXlinker.Device_2_EtherCAT.Term_9_EK1100.Term_10_EK1122.Term_23_EK1100.Term_32_EL2258.MTO_Outputs_10x_Channel_4.Outputs/Output_event_state_1 <-> MTO Outputs 10x Channel 4/Outputs/Output event state 1
//     PlcTask Outputs/GVL_iXlinker.Device_2_EtherCAT.Term_9_EK1100.Term_10_EK1122.Term_23_EK1100.Term_32_EL2258.MTO_Outputs_10x_Channel_4.Outputs/Output_event_state_10 <-> MTO Outputs 10x Channel 4/Outputs/Output event state 10
//     PlcTask Outputs/GVL_iXlinker.Device_2_EtherCAT.Term_9_EK1100.Term_10_EK1122.Term_23_EK1100.Term_32_EL2258.MTO_Outputs_10x_Channel_4.Outputs/Output_event_state_2 <-> MTO Outputs 10x Channel 4/Outputs/Output event state 2
//     PlcTask Outputs/GVL_iXlinker.Device_2_EtherCAT.Term_9_EK1100.Term_10_EK1122.Term_23_EK1100.Term_32_EL2258.MTO_Outputs_10x_Channel_4.Outputs/Output_event_state_3 <-> MTO Outputs 10x Channel 4/Outputs/Output event state 3
//     PlcTask Outputs/GVL_iXlinker.Device_2_EtherCAT.Term_9_EK1100.Term_10_EK1122.Term_23_EK1100.Term_32_EL2258.MTO_Outputs_10x_Channel_4.Outputs/Output_event_state_4 <-> MTO Outputs 10x Channel 4/Outputs/Output event state 4
//     PlcTask Outputs/GVL_iXlinker.Device_2_EtherCAT.Term_9_EK1100.Term_10_EK1122.Term_23_EK1100.Term_32_EL2258.MTO_Outputs_10x_Channel_4.Outputs/Output_event_state_5 <-> MTO Outputs 10x Channel 4/Outputs/Output event state 5
//     PlcTask Outputs/GVL_iXlinker.Device_2_EtherCAT.Term_9_EK1100.Term_10_EK1122.Term_23_EK1100.Term_32_EL2258.MTO_Outputs_10x_Channel_4.Outputs/Output_event_state_6 <-> MTO Outputs 10x Channel 4/Outputs/Output event state 6
//     PlcTask Outputs/GVL_iXlinker.Device_2_EtherCAT.Term_9_EK1100.Term_10_EK1122.Term_23_EK1100.Term_32_EL2258.MTO_Outputs_10x_Channel_4.Outputs/Output_event_state_7 <-> MTO Outputs 10x Channel 4/Outputs/Output event state 7
//     PlcTask Outputs/GVL_iXlinker.Device_2_EtherCAT.Term_9_EK1100.Term_10_EK1122.Term_23_EK1100.Term_32_EL2258.MTO_Outputs_10x_Channel_4.Outputs/Output_event_state_8 <-> MTO Outputs 10x Channel 4/Outputs/Output event state 8
//     PlcTask Outputs/GVL_iXlinker.Device_2_EtherCAT.Term_9_EK1100.Term_10_EK1122.Term_23_EK1100.Term_32_EL2258.MTO_Outputs_10x_Channel_4.Outputs/Output_event_state_9 <-> MTO Outputs 10x Channel 4/Outputs/Output event state 9
//     PlcTask Outputs/GVL_iXlinker.Device_2_EtherCAT.Term_9_EK1100.Term_10_EK1122.Term_23_EK1100.Term_32_EL2258.MTO_Outputs_10x_Channel_5.Outputs/Output_event_state_1 <-> MTO Outputs 10x Channel 5/Outputs/Output event state 1
//     PlcTask Outputs/GVL_iXlinker.Device_2_EtherCAT.Term_9_EK1100.Term_10_EK1122.Term_23_EK1100.Term_32_EL2258.MTO_Outputs_10x_Channel_5.Outputs/Output_event_state_10 <-> MTO Outputs 10x Channel 5/Outputs/Output event state 10
//     PlcTask Outputs/GVL_iXlinker.Device_2_EtherCAT.Term_9_EK1100.Term_10_EK1122.Term_23_EK1100.Term_32_EL2258.MTO_Outputs_10x_Channel_5.Outputs/Output_event_state_2 <-> MTO Outputs 10x Channel 5/Outputs/Output event state 2
//     PlcTask Outputs/GVL_iXlinker.Device_2_EtherCAT.Term_9_EK1100.Term_10_EK1122.Term_23_EK1100.Term_32_EL2258.MTO_Outputs_10x_Channel_5.Outputs/Output_event_state_3 <-> MTO Outputs 10x Channel 5/Outputs/Output event state 3
//     PlcTask Outputs/GVL_iXlinker.Device_2_EtherCAT.Term_9_EK1100.Term_10_EK1122.Term_23_EK1100.Term_32_EL2258.MTO_Outputs_10x_Channel_5.Outputs/Output_event_state_4 <-> MTO Outputs 10x Channel 5/Outputs/Output event state 4
//     PlcTask Outputs/GVL_iXlinker.Device_2_EtherCAT.Term_9_EK1100.Term_10_EK1122.Term_23_EK1100.Term_32_EL2258.MTO_Outputs_10x_Channel_5.Outputs/Output_event_state_5 <-> MTO Outputs 10x Channel 5/Outputs/Output event state 5
//     PlcTask Outputs/GVL_iXlinker.Device_2_EtherCAT.Term_9_EK1100.Term_10_EK1122.Term_23_EK1100.Term_32_EL2258.MTO_Outputs_10x_Channel_5.Outputs/Output_event_state_6 <-> MTO Outputs 10x Channel 5/Outputs/Output event state 6
//     PlcTask Outputs/GVL_iXlinker.Device_2_EtherCAT.Term_9_EK1100.Term_10_EK1122.Term_23_EK1100.Term_32_EL2258.MTO_Outputs_10x_Channel_5.Outputs/Output_event_state_7 <-> MTO Outputs 10x Channel 5/Outputs/Output event state 7
//     PlcTask Outputs/GVL_iXlinker.Device_2_EtherCAT.Term_9_EK1100.Term_10_EK1122.Term_23_EK1100.Term_32_EL2258.MTO_Outputs_10x_Channel_5.Outputs/Output_event_state_8 <-> MTO Outputs 10x Channel 5/Outputs/Output event state 8
//     PlcTask Outputs/GVL_iXlinker.Device_2_EtherCAT.Term_9_EK1100.Term_10_EK1122.Term_23_EK1100.Term_32_EL2258.MTO_Outputs_10x_Channel_5.Outputs/Output_event_state_9 <-> MTO Outputs 10x Channel 5/Outputs/Output event state 9
//     PlcTask Outputs/GVL_iXlinker.Device_2_EtherCAT.Term_9_EK1100.Term_10_EK1122.Term_23_EK1100.Term_32_EL2258.MTO_Outputs_10x_Channel_6.Outputs/Output_event_state_1 <-> MTO Outputs 10x Channel 6/Outputs/Output event state 1
//     PlcTask Outputs/GVL_iXlinker.Device_2_EtherCAT.Term_9_EK1100.Term_10_EK1122.Term_23_EK1100.Term_32_EL2258.MTO_Outputs_10x_Channel_6.Outputs/Output_event_state_10 <-> MTO Outputs 10x Channel 6/Outputs/Output event state 10
//     PlcTask Outputs/GVL_iXlinker.Device_2_EtherCAT.Term_9_EK1100.Term_10_EK1122.Term_23_EK1100.Term_32_EL2258.MTO_Outputs_10x_Channel_6.Outputs/Output_event_state_2 <-> MTO Outputs 10x Channel 6/Outputs/Output event state 2
//     PlcTask Outputs/GVL_iXlinker.Device_2_EtherCAT.Term_9_EK1100.Term_10_EK1122.Term_23_EK1100.Term_32_EL2258.MTO_Outputs_10x_Channel_6.Outputs/Output_event_state_3 <-> MTO Outputs 10x Channel 6/Outputs/Output event state 3
//     PlcTask Outputs/GVL_iXlinker.Device_2_EtherCAT.Term_9_EK1100.Term_10_EK1122.Term_23_EK1100.Term_32_EL2258.MTO_Outputs_10x_Channel_6.Outputs/Output_event_state_4 <-> MTO Outputs 10x Channel 6/Outputs/Output event state 4
//     PlcTask Outputs/GVL_iXlinker.Device_2_EtherCAT.Term_9_EK1100.Term_10_EK1122.Term_23_EK1100.Term_32_EL2258.MTO_Outputs_10x_Channel_6.Outputs/Output_event_state_5 <-> MTO Outputs 10x Channel 6/Outputs/Output event state 5
//     PlcTask Outputs/GVL_iXlinker.Device_2_EtherCAT.Term_9_EK1100.Term_10_EK1122.Term_23_EK1100.Term_32_EL2258.MTO_Outputs_10x_Channel_6.Outputs/Output_event_state_6 <-> MTO Outputs 10x Channel 6/Outputs/Output event state 6
//     PlcTask Outputs/GVL_iXlinker.Device_2_EtherCAT.Term_9_EK1100.Term_10_EK1122.Term_23_EK1100.Term_32_EL2258.MTO_Outputs_10x_Channel_6.Outputs/Output_event_state_7 <-> MTO Outputs 10x Channel 6/Outputs/Output event state 7
//     PlcTask Outputs/GVL_iXlinker.Device_2_EtherCAT.Term_9_EK1100.Term_10_EK1122.Term_23_EK1100.Term_32_EL2258.MTO_Outputs_10x_Channel_6.Outputs/Output_event_state_8 <-> MTO Outputs 10x Channel 6/Outputs/Output event state 8
//     PlcTask Outputs/GVL_iXlinker.Device_2_EtherCAT.Term_9_EK1100.Term_10_EK1122.Term_23_EK1100.Term_32_EL2258.MTO_Outputs_10x_Channel_6.Outputs/Output_event_state_9 <-> MTO Outputs 10x Channel 6/Outputs/Output event state 9
//     PlcTask Outputs/GVL_iXlinker.Device_2_EtherCAT.Term_9_EK1100.Term_10_EK1122.Term_23_EK1100.Term_32_EL2258.MTO_Outputs_10x_Channel_7.Outputs/Output_event_state_1 <-> MTO Outputs 10x Channel 7/Outputs/Output event state 1
//     PlcTask Outputs/GVL_iXlinker.Device_2_EtherCAT.Term_9_EK1100.Term_10_EK1122.Term_23_EK1100.Term_32_EL2258.MTO_Outputs_10x_Channel_7.Outputs/Output_event_state_10 <-> MTO Outputs 10x Channel 7/Outputs/Output event state 10
//     PlcTask Outputs/GVL_iXlinker.Device_2_EtherCAT.Term_9_EK1100.Term_10_EK1122.Term_23_EK1100.Term_32_EL2258.MTO_Outputs_10x_Channel_7.Outputs/Output_event_state_2 <-> MTO Outputs 10x Channel 7/Outputs/Output event state 2
//     PlcTask Outputs/GVL_iXlinker.Device_2_EtherCAT.Term_9_EK1100.Term_10_EK1122.Term_23_EK1100.Term_32_EL2258.MTO_Outputs_10x_Channel_7.Outputs/Output_event_state_3 <-> MTO Outputs 10x Channel 7/Outputs/Output event state 3
//     PlcTask Outputs/GVL_iXlinker.Device_2_EtherCAT.Term_9_EK1100.Term_10_EK1122.Term_23_EK1100.Term_32_EL2258.MTO_Outputs_10x_Channel_7.Outputs/Output_event_state_4 <-> MTO Outputs 10x Channel 7/Outputs/Output event state 4
//     PlcTask Outputs/GVL_iXlinker.Device_2_EtherCAT.Term_9_EK1100.Term_10_EK1122.Term_23_EK1100.Term_32_EL2258.MTO_Outputs_10x_Channel_7.Outputs/Output_event_state_5 <-> MTO Outputs 10x Channel 7/Outputs/Output event state 5
//     PlcTask Outputs/GVL_iXlinker.Device_2_EtherCAT.Term_9_EK1100.Term_10_EK1122.Term_23_EK1100.Term_32_EL2258.MTO_Outputs_10x_Channel_7.Outputs/Output_event_state_6 <-> MTO Outputs 10x Channel 7/Outputs/Output event state 6
//     PlcTask Outputs/GVL_iXlinker.Device_2_EtherCAT.Term_9_EK1100.Term_10_EK1122.Term_23_EK1100.Term_32_EL2258.MTO_Outputs_10x_Channel_7.Outputs/Output_event_state_7 <-> MTO Outputs 10x Channel 7/Outputs/Output event state 7
//     PlcTask Outputs/GVL_iXlinker.Device_2_EtherCAT.Term_9_EK1100.Term_10_EK1122.Term_23_EK1100.Term_32_EL2258.MTO_Outputs_10x_Channel_7.Outputs/Output_event_state_8 <-> MTO Outputs 10x Channel 7/Outputs/Output event state 8
//     PlcTask Outputs/GVL_iXlinker.Device_2_EtherCAT.Term_9_EK1100.Term_10_EK1122.Term_23_EK1100.Term_32_EL2258.MTO_Outputs_10x_Channel_7.Outputs/Output_event_state_9 <-> MTO Outputs 10x Channel 7/Outputs/Output event state 9
//     PlcTask Outputs/GVL_iXlinker.Device_2_EtherCAT.Term_9_EK1100.Term_10_EK1122.Term_23_EK1100.Term_32_EL2258.MTO_Outputs_10x_Channel_8.Outputs/Output_event_state_1 <-> MTO Outputs 10x Channel 8/Outputs/Output event state 1
//     PlcTask Outputs/GVL_iXlinker.Device_2_EtherCAT.Term_9_EK1100.Term_10_EK1122.Term_23_EK1100.Term_32_EL2258.MTO_Outputs_10x_Channel_8.Outputs/Output_event_state_10 <-> MTO Outputs 10x Channel 8/Outputs/Output event state 10
//     PlcTask Outputs/GVL_iXlinker.Device_2_EtherCAT.Term_9_EK1100.Term_10_EK1122.Term_23_EK1100.Term_32_EL2258.MTO_Outputs_10x_Channel_8.Outputs/Output_event_state_2 <-> MTO Outputs 10x Channel 8/Outputs/Output event state 2
//     PlcTask Outputs/GVL_iXlinker.Device_2_EtherCAT.Term_9_EK1100.Term_10_EK1122.Term_23_EK1100.Term_32_EL2258.MTO_Outputs_10x_Channel_8.Outputs/Output_event_state_3 <-> MTO Outputs 10x Channel 8/Outputs/Output event state 3
//     PlcTask Outputs/GVL_iXlinker.Device_2_EtherCAT.Term_9_EK1100.Term_10_EK1122.Term_23_EK1100.Term_32_EL2258.MTO_Outputs_10x_Channel_8.Outputs/Output_event_state_4 <-> MTO Outputs 10x Channel 8/Outputs/Output event state 4
//     PlcTask Outputs/GVL_iXlinker.Device_2_EtherCAT.Term_9_EK1100.Term_10_EK1122.Term_23_EK1100.Term_32_EL2258.MTO_Outputs_10x_Channel_8.Outputs/Output_event_state_5 <-> MTO Outputs 10x Channel 8/Outputs/Output event state 5
//     PlcTask Outputs/GVL_iXlinker.Device_2_EtherCAT.Term_9_EK1100.Term_10_EK1122.Term_23_EK1100.Term_32_EL2258.MTO_Outputs_10x_Channel_8.Outputs/Output_event_state_6 <-> MTO Outputs 10x Channel 8/Outputs/Output event state 6
//     PlcTask Outputs/GVL_iXlinker.Device_2_EtherCAT.Term_9_EK1100.Term_10_EK1122.Term_23_EK1100.Term_32_EL2258.MTO_Outputs_10x_Channel_8.Outputs/Output_event_state_7 <-> MTO Outputs 10x Channel 8/Outputs/Output event state 7
//     PlcTask Outputs/GVL_iXlinker.Device_2_EtherCAT.Term_9_EK1100.Term_10_EK1122.Term_23_EK1100.Term_32_EL2258.MTO_Outputs_10x_Channel_8.Outputs/Output_event_state_8 <-> MTO Outputs 10x Channel 8/Outputs/Output event state 8
//     PlcTask Outputs/GVL_iXlinker.Device_2_EtherCAT.Term_9_EK1100.Term_10_EK1122.Term_23_EK1100.Term_32_EL2258.MTO_Outputs_10x_Channel_8.Outputs/Output_event_state_9 <-> MTO Outputs 10x Channel 8/Outputs/Output event state 9
//   TcoIoTests/TcoIoTests Instance <-> Device 2 (EtherCAT)/Term 9 (EK1100)/Term 10 (EK1122)/Term 23 (EK1100)/Term 33 (EL3164)
//     PlcTask Inputs/GVL_iXlinker.Device_2_EtherCAT.Term_9_EK1100.Term_10_EK1122.Term_23_EK1100.Term_33_EL3164.AI_Standard_Channel_{1..4}.Status/Error <-> AI Standard Channel {1..4}/Status/Error  (4 links)
//     PlcTask Inputs/GVL_iXlinker.Device_2_EtherCAT.Term_9_EK1100.Term_10_EK1122.Term_23_EK1100.Term_33_EL3164.AI_Standard_Channel_1.Status/Limit_1 <-> AI Standard Channel 1/Status/Limit 1
//     PlcTask Inputs/GVL_iXlinker.Device_2_EtherCAT.Term_9_EK1100.Term_10_EK1122.Term_23_EK1100.Term_33_EL3164.AI_Standard_Channel_1.Status/Limit_2 <-> AI Standard Channel 1/Status/Limit 2
//     PlcTask Inputs/GVL_iXlinker.Device_2_EtherCAT.Term_9_EK1100.Term_10_EK1122.Term_23_EK1100.Term_33_EL3164.AI_Standard_Channel_2.Status/Limit_1 <-> AI Standard Channel 2/Status/Limit 1
//     PlcTask Inputs/GVL_iXlinker.Device_2_EtherCAT.Term_9_EK1100.Term_10_EK1122.Term_23_EK1100.Term_33_EL3164.AI_Standard_Channel_2.Status/Limit_2 <-> AI Standard Channel 2/Status/Limit 2
//     PlcTask Inputs/GVL_iXlinker.Device_2_EtherCAT.Term_9_EK1100.Term_10_EK1122.Term_23_EK1100.Term_33_EL3164.AI_Standard_Channel_3.Status/Limit_1 <-> AI Standard Channel 3/Status/Limit 1
//     PlcTask Inputs/GVL_iXlinker.Device_2_EtherCAT.Term_9_EK1100.Term_10_EK1122.Term_23_EK1100.Term_33_EL3164.AI_Standard_Channel_3.Status/Limit_2 <-> AI Standard Channel 3/Status/Limit 2
//     PlcTask Inputs/GVL_iXlinker.Device_2_EtherCAT.Term_9_EK1100.Term_10_EK1122.Term_23_EK1100.Term_33_EL3164.AI_Standard_Channel_4.Status/Limit_1 <-> AI Standard Channel 4/Status/Limit 1
//     PlcTask Inputs/GVL_iXlinker.Device_2_EtherCAT.Term_9_EK1100.Term_10_EK1122.Term_23_EK1100.Term_33_EL3164.AI_Standard_Channel_4.Status/Limit_2 <-> AI Standard Channel 4/Status/Limit 2
//     PlcTask Inputs/GVL_iXlinker.Device_2_EtherCAT.Term_9_EK1100.Term_10_EK1122.Term_23_EK1100.Term_33_EL3164.AI_Standard_Channel_{1..4}.Status/Overrange <-> AI Standard Channel {1..4}/Status/Overrange  (4 links)
//     PlcTask Inputs/GVL_iXlinker.Device_2_EtherCAT.Term_9_EK1100.Term_10_EK1122.Term_23_EK1100.Term_33_EL3164.AI_Standard_Channel_{1..4}.Status/Sync_error <-> AI Standard Channel {1..4}/Status/Sync error  (4 links)
//     PlcTask Inputs/GVL_iXlinker.Device_2_EtherCAT.Term_9_EK1100.Term_10_EK1122.Term_23_EK1100.Term_33_EL3164.AI_Standard_Channel_{1..4}.Status/TxPDO_State <-> AI Standard Channel {1..4}/Status/TxPDO State  (4 links)
//     PlcTask Inputs/GVL_iXlinker.Device_2_EtherCAT.Term_9_EK1100.Term_10_EK1122.Term_23_EK1100.Term_33_EL3164.AI_Standard_Channel_{1..4}.Status/TxPDO_Toggle <-> AI Standard Channel {1..4}/Status/TxPDO Toggle  (4 links)
//     PlcTask Inputs/GVL_iXlinker.Device_2_EtherCAT.Term_9_EK1100.Term_10_EK1122.Term_23_EK1100.Term_33_EL3164.AI_Standard_Channel_{1..4}.Status/Underrange <-> AI Standard Channel {1..4}/Status/Underrange  (4 links)
//     PlcTask Inputs/GVL_iXlinker.Device_2_EtherCAT.Term_9_EK1100.Term_10_EK1122.Term_23_EK1100.Term_33_EL3164.AI_Standard_Channel_{1..4}.Value <-> AI Standard Channel {1..4}/Value  (4 links)
//     PlcTask Inputs/GVL_iXlinker.Device_2_EtherCAT.Term_9_EK1100.Term_10_EK1122.Term_23_EK1100.Term_33_EL3164.InfoData.AdsAddr <-> InfoData/AdsAddr
//     PlcTask Inputs/GVL_iXlinker.Device_2_EtherCAT.Term_9_EK1100.Term_10_EK1122.Term_23_EK1100.Term_33_EL3164.InfoData.State <-> InfoData/State
//     PlcTask Inputs/GVL_iXlinker.Device_2_EtherCAT.Term_9_EK1100.Term_10_EK1122.Term_23_EK1100.Term_33_EL3164.WcState.InputToggle <-> WcState/InputToggle
//     PlcTask Inputs/GVL_iXlinker.Device_2_EtherCAT.Term_9_EK1100.Term_10_EK1122.Term_23_EK1100.Term_33_EL3164.WcState.WcState <-> WcState/WcState
//   TcoIoTests/TcoIoTests Instance <-> Device 2 (EtherCAT)/Term 9 (EK1100)/Term 34 (EL3403)
//     PlcTask Inputs/GVL_iXlinker.Device_2_EtherCAT.Term_9_EK1100.Term_34_EL3403.InfoData.AdsAddr <-> InfoData/AdsAddr
//     PlcTask Inputs/GVL_iXlinker.Device_2_EtherCAT.Term_9_EK1100.Term_34_EL3403.InfoData.State <-> InfoData/State
//     PlcTask Inputs/GVL_iXlinker.Device_2_EtherCAT.Term_9_EK1100.Term_34_EL3403.PM_Inputs_Channel_1.Active_power <-> PM Inputs Channel 1/Active power
//     PlcTask Inputs/GVL_iXlinker.Device_2_EtherCAT.Term_9_EK1100.Term_34_EL3403.PM_Inputs_Channel_2.Active_power <-> PM Inputs Channel 2/Active power
//     PlcTask Inputs/GVL_iXlinker.Device_2_EtherCAT.Term_9_EK1100.Term_34_EL3403.PM_Inputs_Channel_3.Active_power <-> PM Inputs Channel 3/Active power
//     PlcTask Inputs/GVL_iXlinker.Device_2_EtherCAT.Term_9_EK1100.Term_34_EL3403.PM_Inputs_Channel_1.Current <-> PM Inputs Channel 1/Current
//     PlcTask Inputs/GVL_iXlinker.Device_2_EtherCAT.Term_9_EK1100.Term_34_EL3403.PM_Inputs_Channel_2.Current <-> PM Inputs Channel 2/Current
//     PlcTask Inputs/GVL_iXlinker.Device_2_EtherCAT.Term_9_EK1100.Term_34_EL3403.PM_Inputs_Channel_3.Current <-> PM Inputs Channel 3/Current
//     PlcTask Inputs/GVL_iXlinker.Device_2_EtherCAT.Term_9_EK1100.Term_34_EL3403.PM_Inputs_Channel_1.Index <-> PM Inputs Channel 1/Index
//     PlcTask Inputs/GVL_iXlinker.Device_2_EtherCAT.Term_9_EK1100.Term_34_EL3403.PM_Inputs_Channel_2.Index <-> PM Inputs Channel 2/Index
//     PlcTask Inputs/GVL_iXlinker.Device_2_EtherCAT.Term_9_EK1100.Term_34_EL3403.PM_Inputs_Channel_3.Index <-> PM Inputs Channel 3/Index
